(* IEC 61131-3 sources: daoli-st-library/DL_MathData (part 12) *)

(* ---- FC_DL_DintMsToTod.st ---- *)
(*
    FC_DL_DintMsToTod —— 当日毫秒到 TOD 的防御转换
    ------------------------------------------------------------------
    分类      : DL_MathData / TimeConv
    前缀      : FC_DL_
    版本      : 1.0.0
    溯源      : IEC 61131-3 标准 TOD 语义的道莅防御性实现；本件为
                FC_DL_TodToDintMs 的严格逆运算，接口语义由标准定义，
                内部委托平台内建 DINT_TO_TOD，不自行按时基重算；
                外围错误分级、单圈折回、双端钳位与双语文档 100% 自有；
                clean-room 重写，未复制任何闭源厂商源码，参考实现仅限 MIT/Apache 许可
    平台      : 纯 IEC 61131-3，CODESYS V3.5+ / TwinCAT 3 / InoProShop 通用
    作者      : 道莅代码库 · PLC编程专家（R19）
    ------------------------------------------------------------------
    功能说明  : 把「自当日 00:00 起的毫秒数」还原为 TOD，供上层排程件与定时器比较。
                有效域 0~86399999 ms；可接受域 -86400000~172799999 ms（含跨日正负各一圈）。
                核心防御：① 超可接受域直接故障级 031E 早退，绝不对非法值调内建；
                ② 负值按单圈折回当日（先判后算，仅一圈内成立，无循环语句）；
                ③ 钳位只在 0 与 86399999 ms 两端，越界量由 bClampSilently 决定分级；
                ④ 交付门槛：委托 DINT_TO_TOD 内建链，须在 CODESYS / TwinCAT 3 /
                   InoProShop 三平台各编译验证一次（跨平台时间类转换链行为存疑）。
                职责边界：本件只做数值还原，不判时区、不做日历进位。
    错误码    : 16#0001_0400 输入越当日域已被钳位到 0 或 86399999 ms——信息级，正常防御
                16#0001_0401 预留禁用（信息级，不得挪用）
                16#0001_031E 输入超可接受域（< -86400000 ms 或 > 172799999 ms）——故障级，返回 T#0S 且 bValid = FALSE
                16#0001_031F 调用方要求不静默（bClampSilently = FALSE）且发生钳位——故障级，返回钳位值但 bValid = FALSE
                16#0001_0320 预留禁用（故障级，不得挪用）
    码位总账  : 16#0001_0400 用 / 16#0001_0401 预留 ｜ 16#0001_031E 用 / 16#0001_031F 用 / 16#0001_0320 预留
    状态机    : R6 标注 N/A —— 本组件为纯函数无顺序状态机，无 CASE 可写，非法状态不可能出现
    采样约定  : 本件无定时器、无沿检测、无顺序状态；单拍纯计算，结论与任务周期无关。
    修订记录  : 2026-11-16 v1.0.0 首次入库（R19）
*)
FUNCTION FC_DL_DintMsToTod : TOD
VAR_INPUT
    nMsOfDay        : DINT := 0;              // 当日毫秒偏移 [ms]，有效域 0~86399999，可接受域 -86400000~172799999 / day-millisecond offset [ms], valid 0~86399999, accepted -86400000~172799999
    bClampSilently  : BOOL := TRUE;           // TRUE = 越界钳位只置信息码；FALSE = 越界置故障级 / TRUE clamps with info code only, FALSE raises a fault level
END_VAR
VAR_OUTPUT
    eErr            : UDINT;                  // 错误码，0=正常 / error id, 0=ok
    bError          : BOOL;                   // 故障标志，eErr 为故障级时 TRUE / error flag, TRUE on fault-level eErr
    bValid          : BOOL;                   // 返回值是否可用 / return value valid flag
    bClamped        : BOOL;                   // 本拍是否发生钳位 / clamp event in this cycle
END_VAR
VAR CONSTANT
    DL_TOD_MS_MIN   : DINT := 0;              // 当日毫秒下界 [ms] / day-millisecond lower bound [ms]
    DL_TOD_MS_MAX   : DINT := 86399999;       // 当日毫秒上界（24 h − 1 ms） [ms] / day-millisecond upper bound, 24 h minus 1 ms [ms]
    DL_TOD_DAY_MS   : DINT := 86400000;       // 一整天毫秒数（单圈折回用） [ms] / milliseconds of one day, for single-wrap folding [ms]
    DL_TOD_MS_MIN_EXT : DINT := -86400000;    // 可接受下界（跨日回退一圈） [ms] / accepted lower bound, one day backwards [ms]
    DL_TOD_MS_MAX_EXT : DINT := 172799999;    // 可接受上界（跨日超前一圈） [ms] / accepted upper bound, one day forwards [ms]
END_VAR
VAR
    nMs             : DINT;                   // 折回与钳位后的中间毫秒值 [ms] / intermediate millisecond value after folding and clamping [ms]
END_VAR

// 段 1｜返回值与错误状态预置 / segment 1, preset return value and error status
FC_DL_DintMsToTod := T#0S;                    // 故障缺省返回当日零点 / fault default returns midnight
eErr := 0;                                    // 预置无错误 / preset no error
bError := FALSE;                              // 预置无故障 / preset no fault
bValid := FALSE;                              // 预置不可用，通过闸门后置位 / preset invalid, set TRUE after the gates
bClamped := FALSE;                            // 预置未钳位 / preset no clamp

// 段 2｜可接受域闸门（越一圈直接故障级，绝不对非法值调内建）/ segment 2, accepted domain gate
IF (nMsOfDay < DL_TOD_MS_MIN_EXT) OR (nMsOfDay > DL_TOD_MS_MAX_EXT) THEN
    eErr := 16#0001_031E;                     // 超可接受域故障码 / accepted domain exceeded fault id
    bError := TRUE;                           // 置故障标志 / raise the error flag
    bValid := FALSE;                          // 返回值不可用 / return value not usable
    FC_DL_DintMsToTod := T#0S;                // 明确返回零点，不用非法值调内建 / return midnight explicitly, never feed an illegal value to the built-in
    RETURN;                                   // 故障级提前返回 / early return on fault
END_IF

// 段 3｜负值单圈折回当日（先判后算，无循环语句）/ segment 3, fold negative values back by one day
nMs := nMsOfDay;                              // 取入参副本参与运算，不改调用方数据 / copy the input, never modify caller data
IF nMs < DL_TOD_MS_MIN THEN
    nMs := nMs + DL_TOD_DAY_MS;               // 单圈折回：域已由段 2 保证 |nMs| ≤ 一圈 / single wrap is enough, segment 2 bounded the magnitude to one day
END_IF

// 段 4｜当日双端钳位（永不对非法值直接调内建）/ segment 4, clamp on both day bounds
IF nMs < DL_TOD_MS_MIN THEN
    nMs := DL_TOD_MS_MIN;                     // 防御性兜底：折回后仍为负则钳 0 ms / defensive floor, clamp to 0 ms if still negative
    bClamped := TRUE;                         // 记录钳位事件 / record the clamp event
ELSIF nMs > DL_TOD_MS_MAX THEN
    nMs := DL_TOD_MS_MAX;                     // 越上界钳 86399999 ms（24 h − 1 ms） / clamp to 86399999 ms, 24 h minus 1 ms
    bClamped := TRUE;                         // 记录钳位事件 / record the clamp event
END_IF

// 段 5｜钳位分级：静默只置信息码，不静默置故障级但返回钳位值 / segment 5, clamp severity
IF bClamped THEN
    IF bClampSilently THEN
        eErr := 16#0001_0400;                 // 信息级：越当日域已钳位，正常防御，不置故障 / info level, clamped into the day domain, no fault raised
        bValid := TRUE;                       // 钳位值仍可用 / the clamped value is usable
    ELSE
        eErr := 16#0001_031F;                 // 故障级：调用方要求不静默 / fault level, the caller refused silent clamping
        bError := TRUE;                       // 置故障标志 / raise the error flag
        bValid := FALSE;                      // 钳位结果标记为不可用 / the clamped result is flagged unusable
    END_IF
ELSE
    eErr := 0;                                // 一轮内合法输入不进钳位分支 / in-domain input never enters the clamp branch
    bValid := TRUE;                           // 域内结果可用 / in-domain result is usable
END_IF

// 段 6｜委托内建转换（入参已保证落在 0~86399999 ms）/ segment 6, delegate to the built-in conversion
FC_DL_DintMsToTod := DINT_TO_TOD(nMs);        // 委托内建，不自行按时基累加 / delegate to the built-in, never accumulate the time base by hand
END_FUNCTION

(* ---- FC_DL_DintToBcd.st ---- *)
(*
  ==================================================================
  组件名 Component  : FC_DL_DintToBcd
  分类   Category   : DL_MathData
  前缀   Naming     : FC_DL_ ｜ b/n/u/f/t/e/st 类型前缀制（R265）
  码位   Code ID    : 16#0001_0658（故障级）
  版本   Version    : 1.0.0
  复杂度 Complexity  : 低
  功能   Purpose    : DINT → 8 位 BCD（DWORD 容器），负值显式拒绝 + 越域显式拒绝，
                      逐位 MOD 10 / DIV 10 提取后按权装入半字节。
  开源溯源 Origin    : 公开公式 clean-room，参考 BCD 编码公开工程语义（分类与参数域
                      借鉴，零代码复制），本件实现、闸门与码位 100% 自有。
  许可证 License    : MIT
  参考   Reference  : IEC 61131-3:2013 §6.6 算术与移位运算符（MOD / DIV / SHL / OR）
  平台   Platform   : 纯 IEC 61131-3（FOR / MOD / DIV / SHL / OR），三平台通用
  依赖   Depends    : 仅 Standard.library（无库调用）
  分工声明 Split     : FC_DL_ByteToBcd / FC_DL_WordToBcd / FC_DL_UdintToBcd 为既有
                      BCD 编码族（无符号域入口），本件为 DINT 带符号域入口；负值
                      显式拒绝为本件与 UDINT 版本的**行为差异**（写死，禁取绝对值
                      回绕伪装成功）；MOD/DIV 10 原语经派单规格明写授权，本件为
                      BCD 编解码属主；四件互引（R216）。
  归属 Ownership     : 本件无 TYPE 声明；全部引脚为 IEC 标准原生类型。
  ------------------------------------------------------------------
  边界 Boundary     :
                      一 判据顺序（写死）：① nIn < 0 → 故障级码 + udBcd = 0 早退
                         （负值不可 BCD 表示，禁取绝对值回绕）；② nIn > 99999999 →
                         越域故障 + bOvF = TRUE 早退；③ 正常才进入提取；
                      二 两场景一码的反证句（R90）：负值与越域的出口仅 bOvF 一位
                         之差（负值 FALSE / 越域 TRUE），一个输出位即可唯一还原
                         场景，三组以内输出可区分，按 R90 不另立码；
                      三 移位量 4·k（k = 0..7）最大 28 < 32（DWORD 位宽），结构性
                         安全（R48）；
                      四 越域上界常量 DL_BCD_MAX = 99999999 与 8 位 BCD 可表域
                         一致，超域属「不可表」而非「截断后仍可用」，禁静默截断；
                      五 纯函数：无记忆量、无定时器、无边沿实例，每调用重算；
                      六 无全局、无外部变量、无物理地址、无指针。
  错误码 Codes      :
    16#0001_0658【故障级】不可 BCD 编码（nIn < 0 负值，bOvF = FALSE；或
                         nIn > 99999999 越域，bOvF = TRUE）
  码位反证 Note     :
    负值与越域共用一码：出口组合仅 bOvF 一位可区分（边界二反证句），按 R90 不另立。
  验收 Acceptance   :
    算法已证（脚本）：未跑 ｜ 编译器已证（三平台）：未跑
    V1 0 → 16#00000000；V2 99999999 → 16#99999999（恰好整除上界向量）
    V3 -1 → 故障 0658 + bOvF = FALSE + 早退（禁取绝对值）
    V4 100000000 → 故障 0658 + bOvF = TRUE + 早退
    V5 12345678 → 16#12345678
  修订记录 Revision  :
    2026-11-21  v1.0.0  R63 首版（批 1 · 序号 2）
  ==================================================================
*)
FUNCTION FC_DL_DintToBcd : BOOL
VAR_INPUT
    nIn     : DINT := 0; // 待编码整数 [个]，合法域 0..99999999 / the integer to encode, legal from zero to ninety nine million
END_VAR
VAR_OUTPUT
    udBcd   : DWORD := 16#00000000; // 8 位 BCD 输出 [码] / the eight digit BCD output
    bOvF    : BOOL := FALSE;        // 越域标志（仅 nIn > 99999999 置位）[-] / the overflow flag raised only above the BCD domain
    bValid  : BOOL := FALSE;        // 结果可用 [-] / the result usable flag
    eErr    : UDINT := 16#0000_0000; // 错误码，0 = 正常 / the error code, zero is ok
    bError  : BOOL := FALSE;        // 故障标志（故障级码同拍置位，R45 配对）/ the fault flag raised with a fault level code
END_VAR
VAR
    k       : DINT := 0;  // 码元位置索引 [下标]，0..7 / the digit position index from zero to seven
    nShift  : DINT := 0;  // 移位量 [位]，4·k ≤ 28 结构性安全 / the shift amount of four times the position, proven below the word width
    nWork   : DINT := 0;  // 逐位提取工作副本 [个] / the working copy of the digit extraction
    uDig    : USINT := 0; // 当前位码元 [位] / the current digit extracted
END_VAR  // R64 结构补齐：VAR 段缺失的 END_VAR（门禁机械修复）
VAR CONSTANT
    DL_BCD_MAX   : DINT := 99999999;   // 8 位 BCD 可表上界 [个] / the representable ceiling of the eight digit BCD
    DL_BCD_N     : DINT := 8;          // 码元总数 [个] / the digit count of eight
    DL_BCD_TEN   : DINT := 10;         // 十进制提取基数 [个] / the decimal extraction base of ten
    DL_BCD_NIB   : DINT := 4;          // 每码元位宽 [位] / the nibble width of four bits
    DL_BCD_ZERO  : DINT := 0;          // 整型零常量 [个] / the integer zero constant
    DL_BCD_ONE   : DINT := 1;          // 整型一常量 [个] / the integer one constant
END_VAR

// 段 1｜返回值与全部出口预置安全值（R45 四段式第一段）/ segment 1, the preset of the return and every outlet
FC_DL_DintToBcd := FALSE; // 返回值预置假 / preset the return false
udBcd := 16#00000000; // BCD 输出预置全零 [码] / preset the BCD output to all zeros
bOvF := FALSE; // 越域标志预置假 / preset the overflow flag false
bValid := FALSE; // 可用标志预置假 / preset the validity false
eErr := 16#0000_0000; // 错误码预置正常 / preset the code to ok
bError := FALSE; // 故障标志预置假 / preset the error flag false
nWork := DL_BCD_ZERO; // 工作副本预置零 [个] / preset the working copy zero
k := DL_BCD_ZERO; // 索引预置零 / preset the index zero
nShift := DL_BCD_ZERO; // 移位量预置零 [位] / preset the shift amount zero
uDig := 0; // 码元预置零 [位] / preset the digit zero

// 段 2｜判据一：负值显式拒绝（边界一①，禁取绝对值回绕伪装成功）/ segment 2, the negative value rejection
IF nIn < DL_BCD_ZERO THEN // 负值不可 BCD 表示 / a negative value is not representable in BCD
    udBcd := 16#00000000; // 输出强制全零 [码] / force the output to all zeros
    eErr := 16#0001_0658; // 故障级：不可 BCD 编码（负值，bOvF 保持 FALSE 供区分）/ fault grade, not encodable as BCD, the overflow flag stays false for the discrimination
    bError := TRUE; // 同拍置故障标志（R45 配对）/ raise the fault flag on the same scan
    bValid := FALSE; // 结果不可用 / the result is not usable
    RETURN; // 早退 / early return
END_IF

// 段 3｜判据二：越域显式拒绝（边界一②，禁静默截断）/ segment 3, the domain overflow rejection
IF nIn > DL_BCD_MAX THEN // 超 8 位 BCD 可表上界 / above the representable ceiling
    udBcd := 16#00000000; // 输出强制全零 [码] / force the output to all zeros
    bOvF := TRUE; // 置越域标志（与负值场景的唯一区分位）/ raise the overflow flag, the only bit distinguishing this scene
    eErr := 16#0001_0658; // 故障级：不可 BCD 编码（越域）/ fault grade, not encodable as BCD, the domain is exceeded
    bError := TRUE; // 同拍置故障标志（R45 配对）/ raise the fault flag on the same scan
    bValid := FALSE; // 结果不可用 / the result is not usable
    RETURN; // 早退 / early return
END_IF

// 段 4｜逐位提取与按权装入（移位量 4·k ≤ 28 < 32 结构性安全，边界三）/ segment 4, the digit extraction and the weighted packing
nWork := nIn; // 工作副本接管 [个] / take the working copy
FOR k := DL_BCD_ZERO TO DL_BCD_N - DL_BCD_ONE DO // 有界遍历 8 个码元位置 / the bounded traversal over eight digit positions
    uDig := DINT_TO_USINT(nWork MOD DL_BCD_TEN); // 当前位 = nWork MOD 10 [位] / the current digit is the remainder of ten
    nWork := nWork / DL_BCD_TEN; // 副本右移一位（DINT 整除截断，nIn ≥ 0 已证，无负回绕）/ shift the copy one digit right, the truncating division is safe since the input is proven non negative
    nShift := DL_BCD_NIB * k; // 移位量 = 4·k，最大 28 [位] / the shift amount of four times the position
    udBcd := udBcd OR SHL(USINT_TO_DWORD(uDig), nShift); // 码元装入对应半字节（OR 合成）/ pack the digit into its nibble by the or composition
END_FOR

// 段 5｜统一出口 / segment 5, the unified outlet
bValid := TRUE; // 结果可用 / the result is usable
FC_DL_DintToBcd := TRUE; // 返回成功 / return success
END_FUNCTION

(* ---- FC_DL_DintToRealChk.st ---- *)
(*
    FC_DL_DintToRealChk —— DINT 到 REAL 精度告警转换
    ------------------------------------------------------------------
    分类      : DL_MathData / Convert
    前缀      : FC_DL_
    版本      : 1.0.0
    溯源      : IEC 61131-3 标准语义的道莅防御性实现
                （接口语义由 IEC 61131-3 定义，内部委托平台内建 DINT_TO_REAL，
                  外围统一错误码 / 钳位 / 双语文档；clean-room 重写，
                  未复制任何闭源厂商源码，参考实现仅限 MIT/Apache 许可）
    平台      : 纯 IEC 61131-3，CODESYS / TwinCAT / InoProShop 通用
    作者      : 道莅代码库 · PLC编程专家（R17）
    ------------------------------------------------------------------
    功能说明  : 将 DINT 防御性转换为 REAL 并作为返回值输出，转换委托平台内建 DINT_TO_REAL；
                |nIn| 超过 2^24（16777216，REAL 尾数 24 位可精确表示的整数上界）时，
                值照常转换输出，仅置信息级 16#0001_01FC 提示低位精度损失（bError=FALSE、bValid=TRUE）；
                极值对称性防御：采用双侧比较 nIn > 上界 OR nIn < -上界，
                禁用 ABS(nIn) 单侧比较（对 DINT 最小值无回绕，但保持与 R16 LintToLrealChk 同范式，避免后续升位改造引入回绕）；
                钳位方向：无钳位（信息级仅记录，转换结果为最接近的可表值）。
    错误码    : 16#0001_01FC |nIn| 超 2^24 精度极限，转换值低位可能失真——信息级，正常防御
                16#0001_01FD 预留禁用（信息级，不得挪用）
                16#0001_02E8 预留禁用（故障级，不得挪用）
                16#0001_02E9 预留禁用（故障级，不得挪用）
                16#0001_02EA 预留禁用（故障级，不得挪用）
    状态机    : R6 标注 N/A —— 本组件为纯函数无顺序状态机，无 CASE 可写，非法状态不可能出现，故以本节说明替代 ELSE 兜底
    修订记录  : 2026-11-16 v1.0.0 首次入库（R17）
*)
FUNCTION FC_DL_DintToRealChk : REAL
VAR_INPUT
    nIn : DINT; // 待转换整数值，建议域 ±2147483647 [无量纲] / integer value to convert, suggested domain +/-2147483647 [dimensionless]
END_VAR
VAR_OUTPUT
    eErr   : UDINT; // 错误码，0=正常 / error id, 0=ok
    bError : BOOL;  // 是否出错，eErr 非 0 时为 TRUE / error flag, TRUE when eErr is nonzero
    bValid : BOOL;  // 输出是否有效可用 / output valid flag
END_VAR
VAR CONSTANT
    DL_F24_MAX : DINT := 16777216; // REAL 尾数 24 位可精确表示的整数上界 2^24 [无量纲] / 2^24 exact-integer bound of REAL's 24-bit significand [dimensionless]
    DL_REAL_ZERO : REAL := 0.0;    // 返回值预置零（本件无故障路径，仅作预置约定） [无量纲] / preset zero, no fault path in this component [dimensionless]
END_VAR

// 段 1｜返回值与错误状态预置 / segment 1, preset return value and error status
FC_DL_DintToRealChk := DL_REAL_ZERO; // 预置 0.0（本件无故障级路径，仅作预置约定） [无量纲] / preset 0.0, no fault-level path in this component [dimensionless]
eErr   := 0;     // 预置无错误 / preset no error
bError := FALSE; // 预置无故障（本件无故障级路径） / preset no fault, no fault-level path here
bValid := FALSE; // 预置输出无效，通过精度判定后置位 / preset invalid, set TRUE after the precision check

// 段 2｜24 位尾数精度极限判定与主体转换（末段） / segment 2, 24-bit significand precision check and main conversion (final)
FC_DL_DintToRealChk := DINT_TO_REAL(nIn); // 值照常转换（委托平台内建转换语义），本件只告警不钳位 [无量纲] / convert as-is via the built-in conversion, this component warns but never clamps [dimensionless]
IF (nIn > DL_F24_MAX) OR (nIn < -DL_F24_MAX) THEN // 双侧比较，禁用 ABS 单侧式 [无量纲] / two-sided comparison, single-sided ABS form forbidden [dimensionless]
    eErr := 16#0001_01FC; // 信息级：超 2^24 精度极限，低位可能失真，仅记录不钳位 / info level: beyond the 2^24 precision limit, low bits may lose accuracy, recorded only
ELSE
    eErr := 0;            // 精度域内无告警 / within the precision domain, no notice
END_IF
bError := FALSE; // 信息级精度告警不置故障 / info-level precision notice never raises fault
bValid := TRUE;  // 域内或精度告警输出均有效可用 / in-domain or precision-noticed output is valid
END_FUNCTION

(* ---- FC_DL_DintToStringTrim.st ---- *)
(*
    FC_DL_DintToStringTrim —— DINT 到 STRING 的防御字符串化
    ------------------------------------------------------------------
    分类      : DL_MathData / Convert
    前缀      : FC_DL_
    版本      : 1.0.0
    溯源      : IEC 61131-3 标准语义的道莅防御性实现（DINT → STRING，去前导空格与长度钳位）；
                委托平台内建 DINT_TO_STRING 与标准串函数 LEN / MID / LEFT，本件不重实现格式化内核；
                空格修剪、四步截断样板、目标长度闸、错误分级与码位 100% 自有；
                clean-room 重写，未复制任何闭源厂商源码，参考实现仅限 MIT/Apache 许可
    平台      : 纯 IEC 61131-3，CODESYS V3.5+ / TwinCAT 3 / InoProShop 通用
    作者      : 道莅代码库 · PLC编程专家（R20）
    ------------------------------------------------------------------
    功能说明  : 数值要拼进 CSV 行、报文帧、条码内容、文件名时，必须先字符串化。
                各平台 DINT_TO_STRING 的右对齐习惯不一：有的前置空格补齐到固定宽度，
                有的不留空格。带空格的数值混进 CSV 会多出一列，拼进报文会错位一个字节，
                而这类故障在 PLC 侧完全静默，只有上位机解析时才暴露。
                核心防御：① 逐字符定位首个非空格后一次 MID 截取，杜绝「逐字符拼串」的
                   长度与性能问题（拼串会随长度平方级增长）。
                ② 扫描用定长 FOR（上界 255），禁用 WHILE——串函数异常时 WHILE 会死循环，
                   FOR 上界结构性封顶。
                ③ 截断走四步样板（R37）：先把长度一次锁存 → 与目标宽度比较 →
                   截断标志置位先于任何写入 → 按 bAllowTrunc 分路；不允许截断时返回空串
                   并升故障级，绝不返回半截数值——半截数值形如把 12345 写成 123，
                   上位机会把它当成真实数据。
                ④ uTargetMax 引脚钳位在 1~255：0 长度目标无意义；255 是 STRING 型上限（R49 口径），
                   USINT 类型本身的 255 上界即为其第二道保险。
                职责边界：LREAL 字符串化（含非有限值统一文本）归 FC_DL_LrealToStringTrim；
                串处理九函数归 T0-6 家族；本件只管整型方向。
    编译门槛  : 主路径依赖平台内建 DINT_TO_STRING 与标准串函数 LEN / MID / LEFT。
                DINT_TO_STRING 的返回宽度平台间不同（有 11 字符起的多种取值），
                故本件不假设其宽度，一律按 LEN 实测后处理，必要时再按目标长度钳位。
    错误码    : 16#0001_0426 已修剪前导空格（bTrimmed 可查）——信息级，值可用
                16#0001_0427 发生截断且 bAllowTrunc = TRUE（bTruncated 可查）——信息级，值可用
                16#0001_0357 目标长度非法（uTargetMax = 0，或平台 USINT 上限异常）——故障级，返回空串
                16#0001_0358 需要截断但 bAllowTrunc = FALSE——故障级，返回空串
                16#0001_0359 预留禁用（故障级，不得挪用）
    码位总账  : 16#0001_0426 用 / 16#0001_0427 用 ｜ 16#0001_0357 用 / 16#0001_0358 用 / 16#0001_0359 预留
    状态机    : R6 标注 N/A —— 本组件为纯函数无顺序状态机，无 CASE 可写，非法状态不可能出现
    采样约定  : 本件无定时器、无沿检测、无状态；单拍纯计算，结论与任务周期无关。
    修订记录  : 2026-11-16 v1.0.0 首次入库（R20）
*)
FUNCTION FC_DL_DintToStringTrim : STRING(255)
VAR_INPUT
    nIn              : DINT;                  // 待字符串化的数值 [无量纲]，全域 / value to serialise [dimensionless], full DINT domain
    uTargetMax       : USINT := 31;           // 目标缓冲可用长度 [字符]，1~255 / usable target length [characters], 1 to 255
    bAllowTrunc      : BOOL := FALSE;         // TRUE = 允许截断；FALSE = 需截断即故障 / TRUE allows truncation, FALSE turns it into a fault
END_VAR
VAR_OUTPUT
    eErr             : UDINT;                 // 错误码，0=正常 / error id, 0=ok
    bError           : BOOL;                  // 故障标志，eErr 为故障级时 TRUE / error flag, TRUE on fault-level eErr
    bValid           : BOOL;                  // 返回值是否可用（故障级为 FALSE）/ return usable, FALSE on fault level
    bTrimmed         : BOOL;                  // 修剪了前导空格 / leading blanks were trimmed
    bTruncated       : BOOL;                  // 超目标长度发生截断 / truncation to the target length happened
END_VAR
VAR CONSTANT
    DL_STR_CAP_MAX   : USINT := 255;          // STRING 型长度上限 [字符]，R49 口径 / STRING capacity [characters], per R49
    DL_STR_TARGET_MIN : USINT := 1;           // 目标长度下限 [字符] / target length lower bound [characters]
    DL_STR_SCAN_MAX  : INT := 255;            // 扫描上界 [字符]，与 STRING 上限一致 / scan bound [characters], equals the STRING capacity
    DL_STR_BLANK     : STRING(1) := ' ';      // 单个空格字符，修剪判据 / a single blank used by the trim test
    DL_STR_EMPTY     : STRING(1) := '';       // 空串常量，故障缺省返回 / empty string returned on faults
    DL_INT_ZERO      : INT := 0;              // 整型零常量，避免裸字面量 [字符] / integer zero constant [characters]
    DL_INT_ONE       : INT := 1;              // 整型一常量，首个非空格位置起点 [字符] / integer one constant, first non-blank position [characters]
END_VAR
VAR
    sRaw             : STRING(255);           // 内建字符串化原始结果 / raw result of the built-in conversion
    sTrim            : STRING(255);           // 修剪后的中间串 / intermediate string after the trim
    sOut             : STRING(255);           // 最终输出串 / final output string
    nLen             : INT;                   // 原始串有效长度 [字符] / effective length of the raw string [characters]
    nStart           : INT;                   // 首个非空格位置，1 起始，0 = 全为空格 / first non-blank position, 1-based, 0 means all blanks
    nIdx             : INT;                   // 扫描游标 [字符]，1 起始 / scan cursor [characters], 1-based
    nKept            : INT;                   // 修剪后保留长度，一次锁存 [字符] / retained length, latched exactly once [characters]
    nTarget          : INT;                   // 目标长度，由引脚转出 [字符] / target length derived from the pin [characters]
    bFound           : BOOL;                  // 已找到首个非空格标志 / a first non-blank has been found
END_VAR

// 段 1｜返回值与错误状态预置 / segment 1, preset return value and error status
FC_DL_DintToStringTrim := DL_STR_EMPTY;       // 故障缺省返回空串 / fault default returns an empty string
eErr := 0;                                    // 预置无错误 / preset no error
bError := FALSE;                              // 预置无故障 / preset no fault
bValid := FALSE;                              // 预置不可用，通过闸门后置位 / preset invalid, set TRUE after the gates
bTrimmed := FALSE;                            // 预置未修剪 / preset no trim
bTruncated := FALSE;                          // 预置未截断 / preset no truncation
sOut := DL_STR_EMPTY;                         // 输出串清零 / clear the output string
nKept := DL_INT_ZERO;                         // 保留长度清零 / clear the retained length

// 段 2｜目标长度闸：0 长度目标无意义，先判后算 / segment 2, target length gate
IF uTargetMax < DL_STR_TARGET_MIN THEN
    eErr := 16#0001_0357;                     // 故障级：目标长度非法，返回空串 / fault level, illegal target length, return an empty string
    bError := TRUE;                           // 置故障标志 / raise the error flag
    bValid := FALSE;                          // 返回值不可用 / flag the return as unusable
    RETURN;                                   // 出口，不触碰内建 / exit, the built-in is never touched
END_IF
nTarget := USINT_TO_INT(uTargetMax);          // 目标长度转整型 [字符] / convert the target length into an integer [characters]
IF nTarget > USINT_TO_INT(DL_STR_CAP_MAX) THEN
    nTarget := USINT_TO_INT(DL_STR_CAP_MAX);  // 双保险：按 STRING 上限钳位 [字符] / second line of defence, clamp to the STRING capacity [characters]
END_IF

// 段 3｜主体：委托平台内建字符串化 / segment 3, delegate the built-in conversion
sRaw := DINT_TO_STRING(nIn);                  // 数值 → 原始串（可能含前导空格）/ value to raw string, possibly blank padded

// 段 4｜有效长度一次锁存并钳位 / segment 4, latch the effective length once and clamp it
nLen := LEN(sRaw);                            // 原始串长度 [字符] / raw string length [characters]
IF nLen > DL_STR_SCAN_MAX THEN
    nLen := DL_STR_SCAN_MAX;                  // 超容量按上限钳位 [字符] / clamp to the capacity [characters]
ELSIF nLen < DL_INT_ZERO THEN
    nLen := DL_INT_ZERO;                      // 负长度防御，结构性不可达 [字符] / negative length guard, structurally unreachable [characters]
END_IF

// 段 5｜前导空格修剪：定长 FOR 扫描，禁 WHILE / segment 5, leading blank trim with a bounded FOR loop
nStart := DL_INT_ZERO;                        // 0 表示尚未找到非空格 / zero means no non-blank found yet
bFound := FALSE;                              // 扫描标志预置 / preset the scan flag
FOR nIdx := DL_INT_ONE TO nLen DO
    IF NOT bFound THEN
        IF MID(sRaw, DL_INT_ONE, nIdx) <> DL_STR_BLANK THEN
            nStart := nIdx;                   // 记录首个非空格位置 [字符] / record the first non-blank position [characters]
            bFound := TRUE;                   // 扫描标志置位 / raise the scan flag
        END_IF
    END_IF
END_FOR

IF nStart = DL_INT_ZERO THEN
    sTrim := DL_STR_EMPTY;                    // 全为空格：合法的空结果，不是错误 / all blanks, a legal empty result
ELSE
    sTrim := MID(sRaw, nLen - nStart + DL_INT_ONE, nStart); // 一次截取中间段 / extract the retained segment in one call
    IF nStart > DL_INT_ONE THEN
        bTrimmed := TRUE;                     // 确实修剪了前导空格 / blanks were really trimmed
        eErr := 16#0001_0426;                 // 信息级：已修剪前导空格 / info level, leading blanks were trimmed
    END_IF
END_IF

// 段 6｜四步截断样板（R37）：长度锁存 → 宽度比较 → 标志先置 → 按允许分路 / segment 6, the four-step truncation pattern
nKept := LEN(sTrim);                          // 修剪后长度，一次锁存 [字符] / retained length, latched once [characters]
IF nKept > nTarget THEN
    bTruncated := TRUE;                       // 标志先于任何写入 / the flag precedes every write
    IF bAllowTrunc THEN
        sOut := LEFT(sTrim, nTarget);         // 允许截断：按目标长度截取 / truncation allowed, take the target length
        eErr := 16#0001_0427;                 // 信息级：发生截断，值可用 / info level, truncated, still usable
    ELSE
        eErr := 16#0001_0358;                 // 故障级：需截断但不允许 / fault level, truncation needed but not allowed
        bError := TRUE;                       // 置故障标志 / raise the error flag
        bValid := FALSE;                      // 返回值不可用 / flag the return as unusable
        FC_DL_DintToStringTrim := DL_STR_EMPTY; // 返回空串，绝不返回半截数值 / return an empty string, never a partial number
        RETURN;                               // 出口 / exit
    END_IF
ELSE
    sOut := sTrim;                            // 无需截断，直接采用修剪结果 / no truncation, take the trimmed string
END_IF

// 段 7｜发布结果 / segment 7, publish the result
FC_DL_DintToStringTrim := sOut;               // 输出最终串 / publish the final string
bValid := TRUE;                               // 修剪/截断/直通均可用 / usable in every published path
bError := FALSE;                              // 信息级不置故障（双保险）/ info level never raises a fault, second line of defence
END_FUNCTION

(* ---- FC_DL_DintToUintSat.st ---- *)
(*
    FC_DL_DintToUintSat —— DINT 到 UINT 饱和防御转换
    ------------------------------------------------------------------
    分类      : DL_MathData / Convert
    前缀      : FC_DL_
    版本      : 1.0.0
    溯源      : IEC 61131-3 标准语义的道莅防御性实现
                （内部委托平台内建函数，外围统一错误码/钳位/双语文档；
                  未复制任何闭源厂商源码，参考实现仅限 MIT/Apache 许可）
    平台      : 纯 IEC 61131-3，CODESYS / TwinCAT / InoProShop 通用
    作者      : 道莅代码库 · PLC编程专家（R16）
    ------------------------------------------------------------------
    功能说明  : 将 DINT 输入防御性转换为 UINT 并作为返回值输出；
                nIn < 0 时钳位至 0，置信息级 16#0001_01CA（UINT 无符号，负值不可表）；
                nIn 超出 UINT 上界 65535 时钳位至上界，置信息级 16#0001_01CB；
                钳位方向：下界 0 / 上界 65535（双侧饱和）；
                纯整数域输入不存在 NaN/±INF 非有限态，亦无除法运算，故本组件无故障级路径；
                域内转换委托平台内建 DINT_TO_UINT 语义，不重实现数学内核；
                信息级码属正常防御：bError=FALSE、bValid=TRUE，输出钳位后防御值。
    错误码    : 16#0001_01CA 负值输入，已钳位至 0——信息级，正常防御
                16#0001_01CB 输入超 UINT 上界，已钳位至 65535——信息级，正常防御
                16#0001_029D 预留禁用（故障级，不得挪用）
                16#0001_029E 预留禁用（故障级，不得挪用）
                16#0001_029F 预留禁用（故障级，不得挪用）
    状态机    : R6 标注 N/A —— 本组件为纯函数无顺序状态机，无 CASE 可写，非法状态不可能出现，故以本节说明替代 ELSE 兜底
    修订记录  : 2026-11-16 v1.0.0 首次入库（R16）
*)
FUNCTION FC_DL_DintToUintSat : UINT
VAR_INPUT
    nIn : DINT; // 待转换输入 [无量纲] / input value to convert
END_VAR
VAR_OUTPUT
    eErr   : UDINT; // 错误码，0=正常 / error id, 0=ok
    bError : BOOL;  // 是否出错，eErr 非 0 时为 TRUE / error flag, TRUE when eErr is nonzero
    bValid : BOOL;  // 输出是否有效可用 / output valid flag
END_VAR
VAR CONSTANT
    DL_UINT16_MAX : DINT := 65535; // UINT 域上界 65535 [无量纲] / UINT upper bound 65535
END_VAR

// 段 1｜返回值与错误状态预置 / segment 1, preset return value and error status
FC_DL_DintToUintSat := 0; // 故障缺省返回 0 [无量纲] / fault default returns 0
eErr   := 0;     // 预置无错误 / preset no error
bError := FALSE; // 预置无故障（整数域无故障态） / preset no fault (no fault states in integer domain)
bValid := FALSE; // 预置无效，通过钳位判定后置位 / preset invalid, set TRUE after clamp check

// 段 2｜双侧饱和钳位与主体转换（末段） / segment 2, double-side saturating clamp and main conversion (final)
IF nIn < 0 THEN
    FC_DL_DintToUintSat := 0; // 负值钳位至 0（UINT 无符号语义） / negative input clamped to 0 (UINT is unsigned)
    eErr := 16#0001_01CA;     // 信息级：负值已钳零 / info level: negative input clamped to zero
ELSIF nIn > DL_UINT16_MAX THEN
    FC_DL_DintToUintSat := 16#FFFF; // 正向钳位至 UINT 上界 65535 / clamp to UINT upper bound 65535
    eErr := 16#0001_01CB;           // 信息级：超上界已钳位 / info level: above upper bound, clamped
ELSE
    FC_DL_DintToUintSat := DINT_TO_UINT(nIn); // 域内委托平台内建 _TO_ 转换语义 / in-domain delegate to built-in _TO_ conversion
    eErr := 0; // 域内无错误 / in-domain, no error
END_IF
bValid := TRUE; // 域内或钳位输出均有效可用 / in-domain or clamped output is valid
END_FUNCTION

(* ---- FC_DL_DivDintSafeChk.st ---- *)
(*==============================================================================
 * 组件名称 (Component)  : FC_DL_DivDintSafeChk
 * 所属子库 (Sublibrary) : DL_MathData
 * 归属目录 (Directory)  : C:\Library\DL_MathData
 * 当前版本 (Version)    : 1.0.0
 * 分类/来源标签         : 函数（FUNCTION）· 纯函数 · DINT 安全除
 *                         iec-std-wrapper / math-safe
 * 兼容性   (Platform)   : CODESYS 3.5 / TwinCAT 3 / 汇川 InoProShop / 施耐德
 *                         Machine Expert；仅用 IEC 标准 DINT 除法与 MOD 语义
 * 溯源声明 (Provenance) : IEC 61131-3 标准语义的道莅防御性实现——内部委托平台标准库语义，
 *                         外围统一错误码 / 钳位 / 双语注释，严禁重实现数学内核。
 * 功能一句话 (Summary)  : DINT 安全除：除零返回哨兵零并置故障，负最小值除 -1
 *                         的整数溢出显式钳位到 DINT 上限，商余同出可观测。
 *
 * 功能描述 (Function)   : 除零闸先行（除数为零返回哨兵 0 + 故障码）；溢出闸
 *                         拦截 DINT 负最小值除以 -1 的唯一上溢情形，按保守方向
 *                         钳到 DINT 上限；合法路径一次算出商与余数（MOD），
 *                         商余配对输出便于调用方做可逆校验。
 * 与既有件边界 (Boundary): 与 FC_DL_DivLrealSafe 构成整数域/实数域对偶；
 *                         本件哨兵零与「真实商为零」区分靠 bError 与事件码，
 *                         哨兵只出现在故障路径。
 * 码位说明 (Codes)      : 信息 16#0002_304C 整除无余数（余数为零）
 *                         故障 16#0002_304D 除数为零，商返回哨兵零
 *                         故障 16#0002_304E 商溢出（负最小值除 -1），已钳上限
 *                         段 16#02_3_4C~4F 首槽信息级、次槽起故障级。
 * 依赖说明 (Depends)    : 无 DL_ 内部依赖；仅 IEC 标准 DINT 除法 / MOD / 常量。
 * 红线自检 (Redline)    : 零全局依赖 ｜ 零 VAR_EXTERNAL ｜ 零 %I/%Q ｜ 纯 IEC 标准库
 *                         除法前强制判零 ｜ 全变量双语同行注释 ｜ 无定时器实例
 * 修订历史 (Revision)   : 2026-11-18  v1.0.0  首版入库（R32 · 批 2）
 *============================================================================*)

FUNCTION FC_DL_DivDintSafeChk : BOOL
VAR_INPUT
    iDividend : DINT;                   // 被除数 [整数域] / Dividend
    iDivisor  : DINT;                   // 除数 [整数域]，零即触发除零闸 / Divisor, zero triggers the gate
END_VAR
VAR_OUTPUT
    iQuot   : DINT;                     // 商 [整数]，故障路径为哨兵零 / Quotient, sentinel zero on fault
    iRem    : DINT;                     // 余数 [整数]，故障路径为零 / Remainder, zero on fault
    bError  : BOOL;                     // 故障标志，与故障码 304D/304E 配对 / Fault flag paired with codes
    uErrorId: UDINT;                    // 事件码，0 表示无事件 / Event code, zero means none
END_VAR
VAR
    uCode : UDINT;   // 码位暂存，出口单点写入 [码] / Code staging
END_VAR
VAR CONSTANT
    DL_DDS_IMIN : DINT := -2147483648;  // DINT 负最小值 [整数] / DINT most negative value
    DL_DDS_IMAX : DINT := 2147483647;   // DINT 正最大值 [整数] / DINT most positive value
END_VAR

(* 段 1｜输出预置 / Pre-set *)
FC_DL_DivDintSafeChk := FALSE;
iQuot    := 0;
iRem     := 0;
bError   := FALSE;
uErrorId := 16#0000_0000;
uCode    := 16#0000_0000;

(* 段 2｜除零闸：哨兵零 + 故障配对（R45），绝不放行平台异常 / Divide-by-zero gate with sentinel and fault pairing *)
IF iDivisor = 0 THEN
    iQuot    := 0;               // 哨兵零，与真实零商靠 bError 区分 / Sentinel zero, distinguished by bError
    iRem     := 0;
    bError   := TRUE;            // 故障级码配对置位 / Fault flag paired
    uErrorId := 16#0002_304D;    // 故障级：除数为零 / Fault: divisor is zero
    RETURN;
END_IF

(* 段 3｜溢出闸：DINT 负最小值除以 -1 是唯一上溢点，钳到上限 / Overflow gate: the only DINT overflow, clamp to the max *)
IF (iDividend = DL_DDS_IMIN) AND (iDivisor = -1) THEN
    iQuot    := DL_DDS_IMAX;     // 保守方向钳位 / Conservative clamp upward
    iRem     := 0;               // 溢出情形余数无意义，置零 / Remainder meaningless here
    bError   := TRUE;            // 故障级码配对置位 / Fault flag paired
    uErrorId := 16#0002_304E;    // 故障级：商溢出已钳 / Fault: quotient overflow clamped
    FC_DL_DivDintSafeChk := TRUE;
    RETURN;
END_IF

(* 段 4｜合法路径：商余一次算出，余数只判一次 / Legal path: quotient and remainder in one pass *)
iQuot := iDividend / iDivisor;   // 整数除法向零截断（标准语义）/ Integer division truncates toward zero
iRem  := iDividend MOD iDivisor; // 标准取余，符号随被除数 / Standard remainder, sign follows the dividend
IF iRem = 0 THEN
    uCode := 16#0002_304C;       // 信息级：整除无余数 / Info: exact division
END_IF
uErrorId := uCode;               // 码位单点写入 / Single write point
FC_DL_DivDintSafeChk := TRUE;
END_FUNCTION

(* ---- FC_DL_DivLrealSafe.st ---- *)
(*
    组件名称 : FC_DL_DivLrealSafe
    所属子库 : DL_MathData
    当前版本 : 1.0.0
    兼 容 性 : CODESYS V3.5+ / TwinCAT 3 / 汇川 InoProShop；仅依赖 Standard.library
    功能描述 : 浮点防御除法原子，把「除法前置防零」这条红线从散落各件的内联 IF 收成唯一出口。
              取舍 ①：微量分母判故障且不输出伪值 —— 绝不返回 0 冒充有效商，bValid 强制 FALSE，
              逼调用方写分支；返回 0 只会把异常静默带进后面的换算链。
              取舍 ②：溢出判据不用 ABS(商) > LREAL_MAX（商一旦溢出，比较式自身已无意义），
              改用「|分子| / LREAL_MAX > |分母|」等价变形：被除数恒为有限域，除法永不溢出，
              判据结构性安全（R54 预判式内禁乘除溢出的同类纪律）。
              取舍 ③：饱和值与除零分开定性 —— 商超有限域是「可观测的饱和」（bValid TRUE + 信息码），
              分母过小是「无结果」（bValid FALSE + 故障码），两者性质不同，绝不混为一谈。
    开源溯源 : 原创实现，红线手册第六节「除法前置防零」的落地载体；无外部源码参考，码位与分级 100% 自有。；本件为 IEC 61131-3 标准语义的道莅防御性实现（原创实现，零外部源码复制）。
    本文件内含 : FUNCTION FC_DL_DivLrealSafe（单 POU，无配套类型）
    依 赖 : 无 DL_ 内部依赖；Standard.library: 无
    红线自检 : R1 ✓ 零全局变量与外部变量 ｜ R2 ✓ 零物理 IO 地址
              R3 ✓ 纯 IEC 61131-3 ｜ R4 ✓ 微量分母闸 + 阈值合法性闸 + 非有限闸 + 商饱和复检
              R5 ✓ 全变量中英双语同行注释 ｜ R6 N/A 纯函数无顺序状态机，无 CASE 可写
              R7 N/A 无定时器、无沿检测实例 ｜ R8 ✓ 全部阈值常量化
    错误码   : 16#0001_0436 [信息级] 商超有限域已饱和至 ±LREAL_MAX，bValid = TRUE，bError = FALSE
               16#0001_0437 [信息级] 预留禁用（不得挪用）
               16#0001_036F [故障级] |分母| < fDenEps（微量分母），返回 0，bValid = FALSE
               16#0001_0370 [故障级] 阈值参数 fDenEps ≤ 0，返回 0，bValid = FALSE
               16#0001_0371 [故障级] 输入含 NaN 或 ±INF，返回 0，bValid = FALSE
    码位总账 : 16#0001_0436 用 / 16#0001_0437 预留 ｜ 16#0001_036F 用 / 16#0001_0370 用 / 16#0001_0371 用
    遗留假设 : ① NaN 判据用自比较（x = x 为假），±INF 判据用 |x| > LREAL_MAX；两式均为 IEEE 754 语义推导，
              未在 InoProShop 上实测（该平台浮点异常屏蔽字配置未知，若开启 FPU 异常陷阱需先关）。
              ② 商饱和取 ±LREAL_MAX 而非 INF，饱和值可被下游有限性检查捕获，避免 INF 在后续乘法中扩散。
    修订历史 :
        2026-11-16  v1.0.0  首版，R21 批次 1 入库
*)
FUNCTION FC_DL_DivLrealSafe : LREAL
VAR_INPUT
    fNum            : LREAL := 1.0;      // 分子，全域有限实数 [无量纲] / numerator, finite real [dimensionless]
    fDen            : LREAL := 1.0;      // 分母，|fDen| < fDenEps 即判故障 [无量纲] / denominator, a magnitude below fDenEps is a fault [dimensionless]
    fDenEps         : LREAL := 1.0E-12;  // 微量分母阈值，必须 > 0；≤ 0 判故障 [无量纲] / micro denominator threshold, must exceed zero [dimensionless]
END_VAR
VAR_OUTPUT
    eErr            : UDINT;             // 错误码，0=正常；16#0001_04XX 信息级 / 16#0001_03XX 故障级 / error id, 0=ok
    bError          : BOOL;              // 故障级标志，eErr 落 16#0001_03XX 时为 TRUE / fault flag, TRUE on fault-level eErr
    bValid          : BOOL;              // 商是否可用，FALSE 时调用方必须走故障分支 / quotient usable flag, the caller must branch when FALSE
    fRatio          : LREAL;             // 分母安全裕度 = |分母| / fDenEps，≥1 表示远离微量阈，仅调试观察 [倍] / denominator safety margin, debug only [ratio]
END_VAR
VAR
    bNumFin         : BOOL;              // 分子是否有限 / numerator finiteness
    bDenFin         : BOOL;              // 分母是否有限 / denominator finiteness
    bNegResult      : BOOL;              // 商的符号预判，供饱和时取号 / predicted sign of the quotient, used when saturating
    fQuot           : LREAL;             // 商工作寄存器 [无量纲] / quotient working register [dimensionless]
END_VAR
VAR CONSTANT
    DL_DIV_EPS          : LREAL := 1.0E-12;                     // 缺省微量分母阈值 [无量纲] / default micro denominator threshold [dimensionless]
    DL_LREAL_MAX_FINITE : LREAL := 1.7976931348623157E308;      // LREAL 最大有限值，饱和与有限性判据 [无量纲] / largest finite LREAL, saturation and finiteness bound [dimensionless]
    DL_LREAL_ONE        : LREAL := 1.0;                         // 单位哨兵，裕度除法前判分母幅值 [无量纲] / unity sentinel guarding the margin division [dimensionless]
    DL_LREAL_ZERO       : LREAL := 0.0;                         // 零哨兵，避免裸 0 参与比较 [无量纲] / zero sentinel [dimensionless]
    DL_ERR_NONE         : UDINT := 16#0000_0000;                // 无故障 / no error
END_VAR

// 段 1｜返回值与错误状态预置（四段式第一段）/ segment 1, preset the return value and the error state
FC_DL_DivLrealSafe := DL_LREAL_ZERO;    // 故障缺省返回 0 / fault default returns zero
eErr   := DL_ERR_NONE;                  // 预置无错误 / preset no error
bError := FALSE;                        // 预置无故障 / preset no fault
bValid := FALSE;                        // 预置结果不可用 / preset unusable
fRatio := DL_LREAL_ZERO;                // 预置裕度 0 / preset the margin to zero

// 段 2｜阈值合法性闸：阈值本身非法时任何比较都无意义 / segment 2, threshold legality gate
IF fDenEps <= DL_LREAL_ZERO THEN
    eErr   := 16#0001_0370;             // 阈值参数非法（故障级）/ illegal threshold parameter
    bError := TRUE;                     // 置故障标志 / raise the fault flag
    RETURN;                             // 返回 0，bValid 保持 FALSE / return zero, bValid stays FALSE
END_IF

// 段 3｜输入有限性闸：NaN 用自比较，±INF 用幅值越界，两式都必须是显式判据 / segment 3, input finiteness gate
bNumFin := (fNum = fNum) AND (ABS(fNum) <= DL_LREAL_MAX_FINITE);   // 自比较为假即 NaN；幅值越界即 INF / self compare catches NaN, the magnitude bound catches INF
bDenFin := (fDen = fDen) AND (ABS(fDen) <= DL_LREAL_MAX_FINITE);   // 与分子同一判据 / same finite test as for the numerator
IF (NOT bNumFin) OR (NOT bDenFin) THEN
    eErr   := 16#0001_0371;             // 输入非有限（故障级）/ non-finite input, fault level
    bError := TRUE;                     // 置故障标志 / raise the fault flag
    RETURN;                             // 返回 0，bValid 保持 FALSE / return zero, bValid stays FALSE
END_IF

// 段 4｜微量分母闸：域内分母过小一律判故障，不输出伪值 / segment 4, micro denominator gate, never emit a pseudo value
IF ABS(fDen) < fDenEps THEN
    eErr   := 16#0001_036F;             // 微量分母（故障级）/ micro denominator, fault level
    bError := TRUE;                     // 置故障标志 / raise the fault flag
    RETURN;                             // 返回 0，bValid 保持 FALSE；调用方必须走故障分支 / return zero, the caller must branch
END_IF

// 段 5｜分母裕度：|分母| ≤ 1 才做除法，避免调试量自身溢出（R54 口径）/ segment 5, margin computed without any overflowing multiply
IF ABS(fDen) > DL_LREAL_ONE THEN
    fRatio := DL_LREAL_MAX_FINITE;      // 分母远大于阈，裕度封顶表达 / the denominator is far above the threshold, cap the margin
ELSE
    fRatio := ABS(fDen) / fDenEps;      // 分母不超过 1，商不会溢出 / the denominator is at most one, the quotient cannot overflow
END_IF

// 段 6｜商溢出预判：|分子| / LREAL_MAX > |分母| 即商必超有限域，此时禁止直接除 / segment 6, overflow prediction before the division
bNegResult := ((fNum < DL_LREAL_ZERO) AND (fDen > DL_LREAL_ZERO)) OR ((fNum > DL_LREAL_ZERO) AND (fDen < DL_LREAL_ZERO)); // 异号即负商 / unlike signs give a negative quotient
IF (ABS(fNum) / DL_LREAL_MAX_FINITE) > ABS(fDen) THEN
    IF bNegResult THEN
        FC_DL_DivLrealSafe := -DL_LREAL_MAX_FINITE;   // 负向饱和 / saturate negative
    ELSE
        FC_DL_DivLrealSafe := DL_LREAL_MAX_FINITE;    // 正向饱和 / saturate positive
    END_IF
    eErr   := 16#0001_0436;             // 商超有限域已饱和（信息级，不置 bError）/ quotient saturated, info level
    bValid := TRUE;                     // 饱和值可观测，与除零性质不同，结果仍可用 / a saturated value is still observable and usable
    RETURN;                             // 带值返回 / return with the saturated value
END_IF

// 段 7｜域内委托：唯一一次真除法 / segment 7, the single genuine division inside the safe domain
fQuot := fNum / fDen;                   // 分母已过微量闸，商不会发散 / the denominator passed the micro gate, the quotient cannot blow up

// 段 8｜结果复检：预判之外的第二道保险，兜住判据边界误差 / segment 8, result re-check as the second line of defence
IF ABS(fQuot) >= DL_LREAL_MAX_FINITE THEN
    IF bNegResult THEN
        fQuot := -DL_LREAL_MAX_FINITE;  // 负向饱和 / saturate negative
    ELSE
        fQuot := DL_LREAL_MAX_FINITE;   // 正向饱和 / saturate positive
    END_IF
    eErr := 16#0001_0436;               // 商超有限域已饱和（信息级）/ quotient saturated, info level
END_IF

// 段 9｜出口 / segment 9, exit
FC_DL_DivLrealSafe := fQuot;            // 输出商 / publish the quotient
bValid := TRUE;                         // 结果可用 / the result is usable
END_FUNCTION

(* ---- FC_DL_DpFlowSqrtCalc.st ---- *)
// =====================================================================
// FC_DL_DpFlowSqrtCalc.st
// 差压式气体流量换算纯函数 (原名 FC_DL_GasFlowSqrt 因 R148 撞名改为本名)
// Differential-pressure gas flow conversion pure function
// 码位: 16#0001_047B ~ 16#0001_047F (本件独占 5 槽)
// 修改记录: R29 初版 (按 DISPATCH_R29 序 1)
// =====================================================================
FUNCTION FC_DL_DpFlowSqrtCalc : BOOL
VAR_INPUT
    bEnable         : BOOL  := TRUE;      // 使能，FALSE 时输出全 0 / Enable, outputs forced to zero when FALSE
    fDp_Pa          : REAL  := 0.0;       // 实测差压 0~250000 Pa / Measured differential pressure [Pa]
    fKFactor        : REAL  := 1.0;       // 流量系数 0.001~100（含管道/孔板系数）/ Flow coefficient [-]
    fRhoRef_kgm3    : REAL  := 1.2041;    // 参比密度 >0 kg/m³ / Reference density [kg/m3]
    fTRef_C         : REAL  := 20.0;      // 参比温度 -50~200 ℃ / Reference temperature [degC]
    fTNow_C         : REAL  := 20.0;      // 当前温度 -50~200 ℃ / Actual temperature [degC]
    fPRef_kPa       : REAL  := 101.325;   // 参比绝压 >0 kPa / Reference absolute pressure [kPa]
    fPNow_kPa       : REAL  := 101.325;   // 当前绝压 >0 kPa / Actual absolute pressure [kPa]
    fDpMin_Pa       : REAL  := 50.0;      // 开方死区 0~5000 Pa / Square-root dead band [Pa]
    fFlowMax_m3h    : REAL  := 100000.0;  // 量程上限 >0 m³/h / Full-scale flow [m3/h]
END_VAR
VAR_OUTPUT
    fFlow_m3h       : REAL;               // 工况流量 / Actual flow [m3/h]
    fFlowRef_m3h    : REAL;               // 参比工况流量 / Reference flow [m3/h]
    bLowCut         : BOOL;               // 死区截断生效 / Dead-band cut active
    eErr            : UDINT;              // 错误码 / Error code
END_VAR
VAR
    fComp           : REAL;               // 温压补偿因子 sqrt((P/Pref)*(Tref/T)) / Compensation factor [-]
    fTKelvin        : REAL;               // 当前绝对温度（钳下限 1.0 K）/ Actual absolute temperature, clamped [K]
    fTRefKelvin     : REAL;               // 参比绝对温度（钳下限 1.0 K）/ Reference absolute temperature, clamped [K]
    fRhoRatio       : REAL;               // 密度比值 rhoNow/rhoRef / Density ratio [-]
    fRhoNow         : REAL;               // 工况密度估算值 / Estimated actual density [kg/m3]
    fFlowRaw        : REAL;               // 钳制前原始流量 / Raw flow before clamp [m3/h]
    bClamped        : BOOL;               // 量程钳制标志 / Flow clamped to full-scale
END_VAR

// ---------------------------------------------------------------------
// 代码位表（本件独占，勿复用）:
//   16#0001_047B 信息 正常换算完成
//   16#0001_047C 故障 差压 < 0 或任一输入非有限
//   16#0001_047D 故障 参比密度/绝压/温度非法（≤0 或 ≤ -273.15）
//   16#0001_047E 信息 结果超量程已钳制 或 差压落在死区（bLowCut 同拍 TRUE）
//   16#0001_047F 故障 fKFactor ≤ 0 或 fFlowMax_m3h ≤ 0（组态错）
// ---------------------------------------------------------------------

// 默认输出（先清零，故障路径直接返回）
fFlow_m3h    := 0.0;    // 工况流量清零 / Reset actual flow
fFlowRef_m3h := 0.0;    // 参比流量清零 / Reset reference flow
bLowCut      := FALSE;  // 死区标志复位 / Reset dead-band flag
eErr         := 16#0001_047B;  // 预置正常码 / Preset normal code

IF NOT bEnable THEN
    // 使能关闭：输出保持全 0，不置故障级 / Disabled: outputs zero, no fault
    RETURN;  // 直接返回 / Return
END_IF

// ---- 非有限闸（NaN 自反判 + Inf 幅值判，等价 bIsFinite）/ Finite guard ----
IF (fDp_Pa <> fDp_Pa) OR (ABS(fDp_Pa) >= 1.0E12)
   OR (fKFactor <> fKFactor) OR (ABS(fKFactor) >= 1.0E12)
   OR (fRhoRef_kgm3 <> fRhoRef_kgm3) OR (ABS(fRhoRef_kgm3) >= 1.0E12)
   OR (fTRef_C <> fTRef_C) OR (ABS(fTRef_C) >= 1.0E12)
   OR (fTNow_C <> fTNow_C) OR (ABS(fTNow_C) >= 1.0E12)
   OR (fPRef_kPa <> fPRef_kPa) OR (ABS(fPRef_kPa) >= 1.0E12)
   OR (fPNow_kPa <> fPNow_kPa) OR (ABS(fPNow_kPa) >= 1.0E12)
   OR (fDpMin_Pa <> fDpMin_Pa) OR (ABS(fDpMin_Pa) >= 1.0E12)
   OR (fFlowMax_m3h <> fFlowMax_m3h) OR (ABS(fFlowMax_m3h) >= 1.0E12) THEN
    fFlow_m3h    := 0.0;             // 输出走安全侧 / Safe-side output
    fFlowRef_m3h := 0.0;             // 参比输出清零 / Reset reference flow
    eErr         := 16#0001_047C;    // 故障：非有限输入 / Fault: non-finite input
    RETURN;                          // 纯函数不驻留 / Pure function returns
END_IF

// ---- 反接判：差压 < 0 → 故障级，不得取绝对值照算 / Reversed wiring fault ----
IF fDp_Pa < 0.0 THEN
    fFlow_m3h    := 0.0;             // 输出 0 / Zero output
    fFlowRef_m3h := 0.0;             // 参比输出 0 / Zero reference output
    eErr         := 16#0001_047C;    // 故障：差压反接 / Fault: negative dp
    RETURN;                          // 直接返回 / Return
END_IF

// ---- 组态错闸：流量系数与量程 / Configuration fault: K and full scale ----
IF (fKFactor <= 0.0) OR (fFlowMax_m3h <= 0.0) THEN
    fFlow_m3h    := 0.0;             // 输出 0 / Zero output
    fFlowRef_m3h := 0.0;             // 参比输出 0 / Zero reference output
    eErr         := 16#0001_047F;    // 故障：组态错 / Fault: config error
    RETURN;                          // 直接返回 / Return
END_IF

// ---- 参比物性组态错闸 / Reference property configuration fault ----
IF (fRhoRef_kgm3 <= 0.0) OR (fPRef_kPa <= 0.0)
   OR (fTRef_C <= -273.15) OR (fTNow_C <= -273.15) THEN
    fFlow_m3h    := 0.0;             // 输出 0（无状态，不沿用上次值）/ Zero output, no state hold
    fFlowRef_m3h := 0.0;             // 参比输出 0 / Zero reference output
    eErr         := 16#0001_047D;    // 故障：参比物性非法 / Fault: invalid reference property
    RETURN;                          // 直接返回 / Return
END_IF

// ---- 死区判（判在开方前）/ Dead band check before square root ----
IF fDp_Pa <= fDpMin_Pa THEN
    fFlow_m3h    := 0.0;             // 噪声死区截断 / Dead-band cut
    fFlowRef_m3h := 0.0;             // 参比流量同步截断 / Reference flow cut
    bLowCut      := TRUE;            // 截断标志 / Cut active
    eErr         := 16#0001_047E;    // 信息级：死区 / Info: dead band
    RETURN;                          // 直接返回 / Return
END_IF

// ---- 温度转绝对温标，钳下限 1.0 K 防除零 / Convert to K, clamp 1.0 K ----
IF fTNow_C > -272.15 THEN
    fTKelvin := fTNow_C + 273.15;    // 当前温度转 K / Actual temperature to K
ELSE
    fTKelvin := 1.0;                 // 钳下限防除零 / Clamp to 1.0 K
END_IF
IF fTRef_C > -272.15 THEN
    fTRefKelvin := fTRef_C + 273.15; // 参比温度转 K / Reference temperature to K
ELSE
    fTRefKelvin := 1.0;              // 钳下限防除零 / Clamp to 1.0 K
END_IF

// ---- 温压补偿因子 sqrt((P/Pref)*(Tref/T)) / Compensation factor ----
fComp := SQRT((fPNow_kPa / fPRef_kPa) * (fTRefKelvin / fTKelvin));  // 补偿因子 / Compensation factor

// ---- 差压开方 × 流量系数 × 补偿因子 / Square root × K × compensation ----
fFlowRaw := fKFactor * SQRT(fDp_Pa) * fComp;  // 原始工况流量 / Raw actual flow [m3/h]

// ---- 量程钳制（信息级）/ Full-scale clamp (info level) ----
bClamped := FALSE;                       // 钳制标志复位 / Reset clamp flag
IF fFlowRaw > fFlowMax_m3h THEN
    fFlowRaw  := fFlowMax_m3h;           // 钳到量程上限 / Clamp to full scale
    bClamped  := TRUE;                   // 记录钳制 / Mark clamped
END_IF
fFlow_m3h := fFlowRaw;                   // 输出工况流量 / Output actual flow

// ---- 参比流量：fFlow × sqrt(rhoNow/rhoRef) / Reference flow via density ratio ----
fRhoNow := fRhoRef_kgm3 * fComp * fComp; // 由补偿因子反推工况密度 / Actual density from compensation
IF fRhoNow > 0.0 THEN
    fRhoRatio    := fRhoNow / fRhoRef_kgm3;  // 密度比值 / Density ratio [-]
    fFlowRef_m3h := fFlow_m3h * SQRT(fRhoRatio);  // 参比流量 / Reference flow [m3/h]
    IF fFlowRef_m3h > fFlowMax_m3h THEN
        fFlowRef_m3h := fFlowMax_m3h;    // 参比流量同步钳制 / Clamp reference flow
    END_IF
ELSE
    fFlowRef_m3h := fFlow_m3h;           // rhoNow 非法 → 直接复制 / Copy actual flow
    eErr         := 16#0001_047C;        // 槽 2 故障 / Slot 2 fault
    RETURN;                              // 直接返回 / Return
END_IF

// ---- 信息级汇总：钳制优先于正常码 / Info-level aggregation: clamp first ----
IF bClamped THEN
    eErr := 16#0001_047E;                // 信息：超量程钳制 / Info: clamped
END_IF

// 正常完成，返回 TRUE / Normal completion
FC_DL_DpFlowSqrtCalc := TRUE;            // 函数返回值 / Function result

END_FUNCTION

(* ---- FC_DL_DtAddSecondsSat.st ---- *)
(*==============================================================================
 * 组件名称 (Component)  : FC_DL_DtAddSecondsSat
 * 所属子库 (Sublibrary) : DL_MathData
 * 归属目录 (Directory)  : C:\Library\DL_MathData
 * 当前版本 (Version)    : 1.0.0
 * 分类/来源标签         : 函数（FUNCTION）· 纯函数 · 日期时间饱和加法
 *                         iec-std-wrapper / datetime / r81-forward-saturate
 * 兼容性   (Platform)   : CODESYS 3.5 / TwinCAT 3 / 汇川 InoProShop / 施耐德
 *                         Machine Expert；仅用 IEC 标准 DT/TIME 语义与 ABS/TRUNC
 * 溯源声明 (Provenance) : IEC 61131-3 标准语义的道莅防御性实现——内部委托平台标准库语义，
 *                         外围统一错误码 / 钳位 / 双语注释，严禁重实现数学内核。
 * 功能一句话 (Summary)  : 日期时间加秒增量，越域按方向饱和到纪元上下限并报
 *                         故障级（R81 正解方向可饱和），非有限增量提前拦截。
 *
 * 本件存在的意义 (Why this unit exists)：
 *   DT 域加法在跨越纪元上限（库内 DtToDintEpoch 属主的 2038 口径）或下限时，
 *   各平台行为从静默回卷到异常停机不一。本件把「越域」变成显式故障码加饱和值：
 *   正向越界钳到上限、负向越界钳到下限，保守失败方向恒定，调用方看码即知发生了什么。
 *
 * 功能描述 (Function)   : 先对 LREAL 秒增量做非有限双闸（x <> x 判 NaN、
 *                         ABS > 1E308 判 Inf）；零秒恒等返回；增量绝对值超过
 *                         单次 TIME 可表达上限（DL_MAXSEC）时按方向直接饱和；
 *                         合法增量转 TIME 后执行 DT + TIME，结果越上/下限
 *                         同样按方向饱和并报故障码。秒增量按整秒域截断。
 * 与既有件边界 (Boundary): 纪元口径沿用库内 FC_DL_DtToDintEpoch 属主
 *                         （1970-01-01 起、2038-01-19 止的 DINT 秒域）；
 *                         本件只做加法正解方向，不做反解（反解方向按 R81 不饱和）。
 * 码位说明 (Codes)      : 信息 16#0002_3048 零秒增量恒等返回
 *                         故障 16#0002_3049 增量非有限（NaN 或 Inf）
 *                         故障 16#0002_304A 正向越界已饱和到纪元上限
 *                         故障 16#0002_304B 负向越界已饱和到纪元下限
 *                         段 16#02_3_48~4B 首槽信息级、次槽起故障级。
 * 依赖说明 (Depends)    : 无 DL_ 内部依赖；仅 IEC 标准 DT/TIME/ABS/TRUNC 语义。
 * 偏离留档 (Deviation)  : 增量绝对值大于 DL_MAXSEC（24 小时）时不再做精确加法，
 *                         按增量方向直接饱和。理由：单次 TIME 只能表达约 24.8 天，
 *                         且超一天的时间修正必属越域操作，保守方向饱和比跨平台
 *                         回卷行为更安全，此偏离已在头注释与实现双处留档。
 * 红线自检 (Redline)    : 零全局依赖 ｜ 零 VAR_EXTERNAL ｜ 零 %I/%Q ｜ 纯 IEC 标准库
 *                         NaN 用 x <> x、Inf 用 ABS > 1.0E308 精确判据
 *                         全变量双语同行注释 ｜ 无定时器实例 ｜ 无状态机
 * 修订历史 (Revision)   : 2026-11-18  v1.0.0  首版入库（R32 · 批 2）
 *============================================================================*)

FUNCTION FC_DL_DtAddSecondsSat : BOOL
VAR_INPUT
    dtIn     : DT;                       // 基准时刻 [日期时间] / Base date-time
    fSecDelta: LREAL;                    // 秒增量 [s]，整秒域，可为负 / Seconds delta, whole-second domain, may be negative
END_VAR
VAR_OUTPUT
    dtOut    : DT;                       // 结果时刻 [日期时间]，越域时为饱和值 / Result, saturated when out of domain
    bSat     : BOOL;                     // 饱和标志，任一方向越域时为真 / TRUE when saturation happened
    uErrorId : UDINT;                    // 事件码，0 表示无事件 / Event code, zero means none
END_VAR
VAR
    tDelta : TIME;    // 整秒增量转出的时长 [s] / Whole-second delta as a TIME duration
    iSec   : DINT;    // 截断后的整秒增量 [s] / Truncated whole-second delta
    uCode  : UDINT;   // 码位暂存，出口单点写入 [码] / Code staging
END_VAR
VAR CONSTANT
    DL_DAS_MAXSEC  : DINT := 86400;                   // 单次增量上限 [s]，24 小时 / Single delta limit, 24 hours
    DL_DAS_DTMAX   : DT   := DT#2038-01-19-03:14:07;  // 纪元上限，沿用库内 2038 口径 / Epoch upper bound, 2038 convention
    DL_DAS_DTMIN   : DT   := DT#1970-01-01-00:00:00;  // 纪元下限 / Epoch lower bound
END_VAR

(* 段 1｜输出预置 / Pre-set *)
FC_DL_DtAddSecondsSat := FALSE;
dtOut    := dtIn;
bSat     := FALSE;
uErrorId := 16#0000_0000;
uCode    := 16#0000_0000;

(* 段 2｜非有限双闸：NaN 用自反判据，Inf 用实数上限精确判据 / Non-finite gates: NaN by reflexivity, Inf by the real limit *)
IF (fSecDelta <> fSecDelta) OR (ABS(fSecDelta) > 1.0E308) THEN
    uErrorId := 16#0002_3049;    // 故障级：增量非有限，结果保持基准时刻 / Fault: non-finite delta, result stays at base
    RETURN;
END_IF

(* 段 3｜整秒截断：秒域契约，负向同样向零截断 / Whole-second truncation, toward zero in both directions *)
iSec := LREAL_TO_DINT(fSecDelta); // 标准显式转换，向零截断 / Standard explicit conversion, truncates toward zero

(* 段 4｜零秒恒等：信息级告知 / Zero delta identity *)
IF iSec = 0 THEN
    uErrorId := 16#0002_3048;    // 信息级：恒等返回 / Info: identity return
    FC_DL_DtAddSecondsSat := TRUE;
    RETURN;
END_IF

(* 段 5｜越域增量按方向饱和（偏离留档见头注释）/ Oversized delta saturates by direction, see the deviation note *)
IF iSec > DL_DAS_MAXSEC THEN
    dtOut := DL_DAS_DTMAX;       // 正向大步进：饱和到上限 / Positive big step: saturate to the max
    bSat  := TRUE;
    uErrorId := 16#0002_304A;    // 故障级：正向饱和 / Fault: saturated upward
    FC_DL_DtAddSecondsSat := TRUE;
    RETURN;
END_IF
IF iSec < -DL_DAS_MAXSEC THEN
    dtOut := DL_DAS_DTMIN;       // 负向大步进：饱和到下限 / Negative big step: saturate to the min
    bSat  := TRUE;
    uErrorId := 16#0002_304B;    // 故障级：负向饱和 / Fault: saturated downward
    FC_DL_DtAddSecondsSat := TRUE;
    RETURN;
END_IF

(* 段 6｜合法增量：DINT 秒转 TIME 后执行标准 DT 加法 / Legal delta: convert to TIME and add *)
tDelta := DINT_TO_TIME(iSec * 1000);             // 秒转毫秒再转 TIME，乘后仍在 TIME 域内 / Seconds to ms to TIME, in range
dtOut  := dtIn + tDelta;                         // 标准 DT + TIME 语义 / Standard DT plus TIME

(* 段 7｜越界检测与方向饱和 / Bound check and directional saturation *)
IF dtOut > DL_DAS_DTMAX THEN
    dtOut := DL_DAS_DTMAX;       // 正向越界：钳上限 / Upward out of bounds: clamp to the max
    bSat  := TRUE;
    uErrorId := 16#0002_304A;    // 故障级：正向饱和 / Fault: saturated upward
ELSIF dtOut < DL_DAS_DTMIN THEN
    dtOut := DL_DAS_DTMIN;       // 负向越界：钳下限 / Downward out of bounds: clamp to the min
    bSat  := TRUE;
    uErrorId := 16#0002_304B;    // 故障级：负向饱和 / Fault: saturated downward
END_IF
FC_DL_DtAddSecondsSat := TRUE;
END_FUNCTION

(* ---- FC_DL_DtToDintEpoch.st ---- *)
(*
    FC_DL_DtToDintEpoch —— DATE_AND_TIME 到 Unix 纪元秒
    ------------------------------------------------------------------
    分类      : DL_MathData / Convert
    前缀      : FC_DL_
    版本      : 1.0.0
    溯源      : IEC 61131-3 标准语义的道莅防御性实现（DATE_AND_TIME → Unix 纪元秒）；
                委托平台内建 DT_TO_DINT 完成秒口径换算，本件不重实现历法内核；
                纪元下域闸门、Y2038 上域饱和出口、错误分级与码位 100% 自有；
                clean-room 重写，未复制任何闭源厂商源码，参考实现仅限 MIT/Apache 许可
    平台      : 纯 IEC 61131-3，CODESYS V3.5+ / TwinCAT 3 / InoProShop 通用
    作者      : 道莅代码库 · PLC编程专家（R20）
    ------------------------------------------------------------------
    功能说明  : 把 PLC 本地时刻统一落成 MES / 日志通用的 Unix 纪元秒（1970-01-01T00:00:00Z 起算）。
                核心防御：① 早于纪元的时刻在类型域上可能出现（平台允许任意 DT 位型），
                   一律在调用内建前拦下——域外调用内建会得到回绕负值，混入日志后无法追溯；
                ② Y2038 是 DINT 秒域硬边界：结果超域时饱和至上限并升故障级，
                   绝不让溢出后的负秒静默流进 MES 台账；
                ③ 结果进入 Y2038 邻近带（2035-01-01 起）只发信息级告警，
                   量仍然可用——告警与故障分级严格分开，HMI 不因提示码停机；
                ④ 负秒重判为第二道防线：域门已保证不可达，仍保留判据，
                   防平台 DT_TO_DINT 在内建层做异常符号处理。
                职责边界：反方向（纪元秒 → DT）归 FC_DL_DintEpochToDt；
                日期天数化归 FC_DL_DateToDintDays；本件只承担「时刻 → 秒」单向标准化。
    编译门槛  : 主路径依赖平台内建 DT_TO_DINT（DT 秒口径），三平台标准库均提供。
                若目标平台缺该内建，按合成路径落地：DT_TO_DATE 取天数、DT_TO_TOD 取当日
                毫秒再折秒，nSec = nDays * DL_SEC_PER_DAY + nSecOfDay；乘法前先判
                nDays < DL_EPOCH_SEC_MAX / DL_SEC_PER_DAY（先判后算，防 DINT 乘法溢出）。
                合成路径不改变本件的闸门顺序与出口，仅替换段 3 的内建调用。
    错误码    : 16#0001_040C Y2038 邻近告警（结果已进入 2035-01-01 起算的告警带）——信息级，值仍可用
                16#0001_040D 预留禁用（信息级，不得挪用）
                16#0001_0330 输入时刻早于纪元（1970-01-01-00:00:00 之前）——故障级，返回 0
                16#0001_0331 结果超出 DINT 秒域（Y2038 2038-01-19T03:14:07Z 之后）——故障级，已饱和至上限
                16#0001_0332 预留禁用（故障级，不得挪用）
    码位总账  : 16#0001_040C 用 / 16#0001_040D 预留 ｜ 16#0001_0330 用 / 16#0001_0331 用 / 16#0001_0332 预留
    状态机    : R6 标注 N/A —— 本组件为纯函数无顺序状态机，无 CASE 可写，非法状态不可能出现
    采样约定  : 本件无定时器、无沿检测、无状态；单拍纯计算，结论与任务周期无关。
    修订记录  : 2026-11-16 v1.0.0 首次入库（R20）
*)
FUNCTION FC_DL_DtToDintEpoch : DINT
VAR_INPUT
    dtIn             : DATE_AND_TIME;         // 输入时刻 [日期时间]，有效域自 1970-01-01-00:00:00 起 / input instant [date and time], domain starts at the epoch
END_VAR
VAR_OUTPUT
    eErr             : UDINT;                 // 错误码，0=正常 / error id, 0=ok
    bError           : BOOL;                  // 故障标志，eErr 为故障级时 TRUE / error flag, TRUE on fault-level eErr
    bValid           : BOOL;                  // 返回值是否可用（故障级为 FALSE）/ return usable, FALSE on fault level
END_VAR
VAR CONSTANT
    DL_EPOCH_SEC_MAX : DINT := 2147483647;    // DINT 秒域上限，即 2038-01-19T03:14:07Z [s] / DINT second domain top, the Y2038 instant [s]
    DL_Y2038_WARN_SEC : DINT := 2051222400;   // Y2038 告警阈值，即 2035-01-01T00:00:00Z [s] / Y2038 warning threshold [s]
    DL_SEC_PER_DAY   : DINT := 86400;         // 每日秒数 [s/日]，合成路径备用量 / seconds per day [s/day], reserved for the synthesis path
    DL_DINT_ZERO     : DINT := 0;             // 有符号零常量，避免裸字面量 [s] / signed zero constant [s]
    DL_EPOCH_DT_ZERO : DATE_AND_TIME := DT#1970-01-01-00:00:00; // 纪元起点时刻 / the epoch instant
END_VAR
VAR
    nSec             : DINT;                  // 纪元秒中间量 [s] / epoch second intermediate [s]
END_VAR

// 段 1｜返回值与错误状态预置 / segment 1, preset return value and error status
FC_DL_DtToDintEpoch := DL_DINT_ZERO;          // 故障缺省返回 0 [s] / fault default returns zero [s]
eErr := 0;                                    // 预置无错误 / preset no error
bError := FALSE;                              // 预置无故障 / preset no fault
bValid := FALSE;                              // 预置不可用，通过闸门后置位 / preset invalid, set TRUE after the gates
nSec := DL_DINT_ZERO;                         // 中间量清零 / clear the intermediate

// 段 2｜下域闸门：早于纪元的时刻在调用内建之前拦下 / segment 2, epoch lower gate precedes any built-in call
IF dtIn < DL_EPOCH_DT_ZERO THEN
    eErr := 16#0001_0330;                     // 故障级：输入早于纪元 / fault level, the input precedes the epoch
    bError := TRUE;                           // 置故障标志 / raise the error flag
    bValid := FALSE;                          // 返回值不可用 / flag the return as unusable
    FC_DL_DtToDintEpoch := DL_DINT_ZERO;      // 确定缺省值 0 / deterministic default of zero
    RETURN;                                   // 出口，不触碰内建 / exit, the built-in is never touched
END_IF

// 段 3｜主体：域内才委托平台内建（秒口径） / segment 3, delegate the built-in only inside the domain
nSec := DT_TO_DINT(dtIn);                     // 内建换算：DT → 纪元秒 [s] / built-in conversion from DT to epoch seconds [s]

// 段 4｜负值第二道防线（域门已保证不可达，保留以防内建层异常符号处理）/ segment 4, second line of defence against a negative result
IF nSec < DL_DINT_ZERO THEN
    eErr := 16#0001_0330;                     // 故障级：内建层给出负秒，等价于早于纪元 / fault level, a negative second means the epoch was underflowed
    bError := TRUE;                           // 置故障标志 / raise the error flag
    bValid := FALSE;                          // 返回值不可用 / flag the return as unusable
    FC_DL_DtToDintEpoch := DL_DINT_ZERO;      // 确定缺省值 0 / deterministic default of zero
    RETURN;                                   // 出口 / exit
END_IF

// 段 5｜Y2038 上域闸：溢出不容静默，饱和并升故障级 / segment 5, Y2038 upper gate, saturation is reported as a fault
IF nSec > DL_EPOCH_SEC_MAX THEN
    nSec := DL_EPOCH_SEC_MAX;                 // 饱和至 DINT 秒域上限 [s] / saturate to the DINT second domain top [s]
    FC_DL_DtToDintEpoch := nSec;              // 发布饱和值供 HMI 观察 / publish the saturated value so HMI can see the overrun
    eErr := 16#0001_0331;                     // 故障级：结果超 DINT 秒域，已饱和 / fault level, the result passed the domain and was saturated
    bError := TRUE;                           // 置故障标志 / raise the error flag
    bValid := FALSE;                          // 饱和值不可用于台账 / the saturated value must not enter the ledgers
    RETURN;                                   // 出口 / exit
END_IF

// 段 6｜发布结果与 Y2038 邻近告警（信息级永不置 bError）/ segment 6, publish and raise the info-level Y2038 warning
FC_DL_DtToDintEpoch := nSec;                  // 输出纪元秒 [s] / publish the epoch seconds [s]
bValid := TRUE;                               // 域内与告警带内均可用 / usable inside the domain and inside the warning band
IF nSec >= DL_Y2038_WARN_SEC THEN
    eErr := 16#0001_040C;                     // 信息级：Y2038 邻近告警，值仍可用 / info level, near Y2038, the value is still usable
END_IF
END_FUNCTION

(* ---- FC_DL_DtToTodWrap.st ---- *)
(*
  ==================================================================
  组件名 Component  : FC_DL_DtToTodWrap
  分类   Category   : DL_MathData
  前缀   Naming     : FC_DL_ ｜ b/n/u/f/t/e/st 类型前缀制（R265）
  码位   Code ID    : 16#0001_0652（信息级）
  版本   Version    : 1.0.0
  复杂度 Complexity  : 低
  功能   Purpose    : 从 DT 提取当日秒数（0..86399）与 TOD，日模 86400 显式化。
  开源溯源 Origin    : IEC 61131-3 标准语义的道莅防御性实现（clean-room，无第三方代码行）
  许可证 License    : MIT
  参考   Reference  : IEC 61131-3:2013 §6.4.3 日期时间类型（DT / TOD）与 §6.5.1 时长域语义
  平台   Platform   : 纯 IEC 61131-3（MOD / 委托 / TOD 类型），三平台通用
  依赖   Depends    : FC_DL_DtToDintEpoch（时刻→纪元秒属主，其内部委托 FC_DL_DateToDintDays
                      完成天序数换算）；FC_DL_DintMsToTod（毫秒→TOD 还原属主）。
                      本件全程委托，不内联任何历法算法（R140 / R216）。
  分工声明 Split     : FC_DL_TodAddWrap / FC_DL_TodDiffWrap 为 TOD 运算属主；
                      FC_DL_TimeToDintMs 为 TIME 域属主；FC_DL_DtToDintEpoch 为绝对纪元秒属主；
                      本件为「DT → 当日秒 / TOD 提取」，四件边界写死（R216 双向互引）。
  归属 Ownership     : 本件无 TYPE 声明；引用件的码位随其属主回传（R66）。
  编译门槛 Gate      : 交付门槛：主路径委托 FC_DL_DtToDintEpoch（其内含 DT_TO_DINT 内建链）
                      与 FC_DL_DintMsToTod（内含 DINT_TO_TOD 内建链），须在 CODESYS /
                      TwinCAT 3 / InoProShop 三平台各编译验证一次（R64）。
  ------------------------------------------------------------------
  边界 Boundary     :
                      一 基准无效闸：dtIn 早于 DT#1970-01-01-00:00:00 视为未初始化或非法
                         时间戳，返回哨兵零点 + 信息级码 + bValid = FALSE，禁止把负天数
                         MOD 成一个看似合法的时刻（还原方向不饱和，R81：返回哨兵零点）；
                      二 日模 86400 显式化：diSecOfDay = ((纪元秒 MOD 86400) + 86400) MOD 86400，
                         双 MOD 保证负数路径也不落到负值域（域外不可达，证明在注释内）；
                      三 todOut 经 FC_DL_DintMsToTod 还原（毫秒域 × 1000），不自行拼 TOD 位型；
                      四 委托件的返回值与 bValid 由两个独立变量承接（R62-D5 教训：禁双写）；
                      五 纯函数：无记忆量、无定时器、无边沿实例，每调用重算。
  错误码 Codes      :
    16#0001_0652【信息级】输入时刻早于纪元基准，已返哨兵零点（bValid = FALSE，不置 bError）
    委托件故障码（16#0001_0330 / 0331 等）按「码随属主」原样回传（R66），本件不另立码。
  码位反证 Note     :
    本件唯一自有码 0652 不可省略：「早于基准」与「委托件进位失败」在出口上都是 bValid = FALSE
    且 todOut = 零点，但两者的处置主体与责任方不同（调用方时间戳未初始化 vs 平台位型承载异常），
    合并会让现场把「未初始化」误判为平台缺陷（R90 反证句）。
  验收 Acceptance   :
    算法已证（脚本）：未跑 ｜ 编译器已证（三平台）：未跑
    V1 DT#1970-01-01-00:00:00 → 0 秒、todOut = 00:00:00、bValid = TRUE
    V2 DT#2024-02-29-23:59:59 → 86399 秒（闰日不计日差，只取当日秒）
    V3 DT#2024-03-01-00:00:00 → 0 秒（日推进不残留）
    V4 DT#1970-01-01-00:00:00 之前的时刻 → bValid = FALSE + 码 0652 + 哨兵零点
    V5 DT#2106-02-07-06:28:15 → 23295 秒（6×3600 + 28×60 + 15，当日秒，跨 32 位不溢出）
    V6 DT#1970-01-02-00:00:00 → 0 秒（日推进归零）
  修订记录 Revision  :
    2026-11-21  v1.0.0  R62 首版（批 3 · 序号 7）
  ==================================================================
*)
FUNCTION FC_DL_DtToTodWrap : BOOL
VAR_INPUT
    dtIn : DT := DT#1970-01-01-00:00:00; // 输入时刻 [日期时间]，有效域自 1970-01-01-00:00:00 起 / the input instant, the domain starts at the epoch
END_VAR
VAR_OUTPUT
    todOut     : TOD;   // 当日时刻 [时刻]，00:00:00 ~ 23:59:59 / the time of day
    diSecOfDay : DINT;  // 当日秒数 [秒]，0..86399 / the second of the day
    bValid     : BOOL;  // 输出可用（早于基准与委托故障为 FALSE）[-] / the output is usable
    eErr       : UDINT; // 错误码，0 = 正常 / the error code, zero is ok
    bError     : BOOL;  // 故障标志，故障级码同拍置位（R45 配对）；信息级恒 FALSE / the fault flag, raised with a fault level code only
END_VAR
VAR
    _nEpochSec   : DINT := 0;                // 委托返回的纪元秒 [秒] / the epoch second returned by the delegate
    _bEpochValid : BOOL := FALSE;            // 委托 bValid 承接量（独立承接，禁双写）/ the delegate valid holder, never double written
    _bEpochErr   : BOOL := FALSE;            // 委托 bError 承接量（独立承接）/ the delegate fault holder, never double written
    _uEpochErr   : UDINT := 16#0000_0000;    // 委托错误码承接量 [码] / the delegate error code holder
    _nMsOfDay    : DINT := 0;                // 当日毫秒偏移 [毫秒] / the millisecond offset inside the day
    _todWork     : TOD := TOD#00:00:00;      // 委托 TOD 返回值承接量 [时刻] / the delegate time of day holder
    _bTodValid   : BOOL := FALSE;            // 委托 TOD 可用位承接量 / the delegate time of day usable holder
    _bTodErr     : BOOL := FALSE;            // 委托 TOD 故障位承接量 / the delegate time of day fault holder
    _uTodErr     : UDINT := 16#0000_0000;    // 委托 TOD 错误码承接量 [码] / the delegate time of day error code holder
    _bTodClamped : BOOL := FALSE;            // 委托 TOD 钳位位承接量（仅留档，不参与分级）/ the delegate clamp holder, recorded only
END_VAR  // R64 结构补齐：VAR 段缺失的 END_VAR（门禁机械修复）
VAR CONSTANT
    DL_DTT_SEC_PER_DAY : DINT := 86400;      // 每日秒数（日模）[秒] / the seconds of one day, the day modulus
    DL_DTT_MS_PER_SEC : DINT := 1000;        // 每秒毫秒数（毫秒域换算）[毫秒] / the milliseconds of one second
    DL_DTT_DINT_ZERO : DINT := 0;             // 整型零常量 [秒] / the integer zero constant
    DL_DTT_TOD_ZERO : TOD := TOD#00:00:00;   // 时刻哨兵零点 [时刻] / the sentinel midnight
    DL_DTT_EPOCH : DT := DT#1970-01-01-00:00:00; // 纪元基准时刻 [日期时间] / the epoch baseline instant
END_VAR

// 段 1｜返回值与全部出口预置安全值（R45 四段式第一段）/ segment 1, preset every outlet to its safe value
FC_DL_DtToTodWrap := FALSE; // 返回值预置假 / preset the return false
todOut := DL_DTT_TOD_ZERO; // 时刻预置哨兵零点 [时刻] / preset the sentinel midnight
diSecOfDay := DL_DTT_DINT_ZERO; // 当日秒数预置零 [秒] / preset the second of the day zero
bValid := FALSE; // 可用标志预置假，过闸后置位 / preset the validity false, raised after the gates
eErr := 16#0000_0000; // 错误码预置正常 / preset the code to ok
bError := FALSE; // 故障标志预置假 / preset the fault flag false
_nEpochSec := DL_DTT_DINT_ZERO; // 纪元秒承接量清零 [秒] / clear the epoch second holder
_bEpochValid := FALSE; // 委托可用位承接量清零 / clear the delegate usable holder
_bEpochErr := FALSE; // 委托故障位承接量清零 / clear the delegate fault holder
_uEpochErr := 16#0000_0000; // 委托码承接量清零 [码] / clear the delegate code holder
_nMsOfDay := DL_DTT_DINT_ZERO; // 当日毫秒清零 [毫秒] / clear the millisecond offset
_todWork := DL_DTT_TOD_ZERO; // 时刻承接量清零 [时刻] / clear the time of day holder
_bTodValid := FALSE; // 委托 TOD 可用位清零 / clear the time of day usable holder
_bTodErr := FALSE; // 委托 TOD 故障位清零 / clear the time of day fault holder
_uTodErr := 16#0000_0000; // 委托 TOD 码清零 [码] / clear the time of day code
_bTodClamped := FALSE; // 委托钳位位清零 / clear the delegate clamp holder

// 段 2｜基准无效闸：早于纪元的时刻不交给委托件（边界一，还原方向不饱和，R81）/ segment 2, the epoch baseline gate
IF dtIn < DL_DTT_EPOCH THEN // 未初始化或非法时间戳 / an uninitialised or illegal timestamp
    todOut := DL_DTT_TOD_ZERO; // 哨兵零点 [时刻] / the sentinel midnight
    diSecOfDay := DL_DTT_DINT_ZERO; // 哨兵零秒 [秒] / the sentinel zero second
    bValid := FALSE; // 输出不可用 / the output is not usable
    eErr := 16#0001_0652; // 信息级：输入早于纪元基准 / informational, the input precedes the epoch baseline
    bError := FALSE; // 明确不置故障标志（信息级，R285）/ keep the fault flag false, this is informational
    RETURN; // 早退，绝不把负天数交给委托件 / early return, a negative day count never reaches the delegate
END_IF

// 段 3｜委托时刻→纪元秒（R140 委托优先；返回值与可用位分承）/ segment 3, delegate the instant to the epoch second
_nEpochSec := FC_DL_DtToDintEpoch(dtIn := dtIn, eErr => _uEpochErr, bError => _bEpochErr, bValid => _bEpochValid); // 委托纪元秒换算 [秒] / delegate the epoch conversion
IF (NOT _bEpochValid) OR _bEpochErr THEN // 委托失败：码随属主回传（R66）/ the delegate failed, the code follows its owner
    eErr := _uEpochErr; // 原样回传委托码 [码] / replay the delegate code as is
    bError := _bEpochErr; // 原样回传委托故障位 / replay the delegate fault bit as is
    bValid := FALSE; // 输出不可用 / the output is not usable
    todOut := DL_DTT_TOD_ZERO; // 哨兵零点 [时刻] / the sentinel midnight
    diSecOfDay := DL_DTT_DINT_ZERO; // 哨兵零秒 [秒] / the sentinel zero second
    RETURN; // 早退 / early return
END_IF

// 段 4｜日模 86400 抽取当日秒（边界二：双 MOD 保证任何输入都落 0..86399）/ segment 4, the day modulus extraction
// 域外不可达证明：段 2 已证 dtIn ≥ 纪元，委托件已证返回值非负，故首层 MOD 的结果已在 [0, 86399]；
// 第二次「+ 86400 再 MOD」为结构对称的二重防御，保证任何未来改动都不会引入负值域出口。
// domain proof: the gate above guarantees a non negative epoch second, so the first modulus already lands inside the day;
// the second fold is a structural second line of defence against any future refactor.
diSecOfDay := ((_nEpochSec MOD DL_DTT_SEC_PER_DAY) + DL_DTT_SEC_PER_DAY) MOD DL_DTT_SEC_PER_DAY; // 当日秒数 [秒] / the second of the day

// 段 5｜委托毫秒→TOD 还原（边界三：不自行拼 TOD 位型）/ segment 5, delegate the millisecond offset back to a time of day
_nMsOfDay := diSecOfDay * DL_DTT_MS_PER_SEC; // 当日毫秒偏移（上界 86399000，DINT 内不溢出）[毫秒] / the millisecond offset, bounded by eighty six million four hundred thousand
_todWork := FC_DL_DintMsToTod(nMsOfDay := _nMsOfDay, bClampSilently := TRUE, eErr => _uTodErr, bError => _bTodErr, bValid => _bTodValid, bClamped => _bTodClamped); // 委托还原 [时刻] / delegate the restoration
IF (NOT _bTodValid) OR _bTodErr THEN // 委托失败：码随属主回传 / the delegate failed, the code follows its owner
    eErr := _uTodErr; // 原样回传委托码 [码] / replay the delegate code as is
    bError := _bTodErr; // 原样回传委托故障位 / replay the delegate fault bit as is
    bValid := FALSE; // 输出不可用 / the output is not usable
    todOut := DL_DTT_TOD_ZERO; // 哨兵零点 [时刻] / the sentinel midnight
    RETURN; // 早退 / early return
END_IF

// 段 6｜统一出口 / segment 6, the unified outlet
todOut := _todWork; // 时刻出口 [时刻] / the time of day outlet
bValid := TRUE; // 域内输出可用 / the in-domain output is usable
FC_DL_DtToTodWrap := TRUE; // 返回成功 / return success
END_FUNCTION

(* ---- FC_DL_DwordToHexString.st ---- *)
(*
    组件名称 : FC_DL_DwordToHexString
    所属子库 : DL_MathData
    当前版本 : 1.0.0
    兼 容 性 : CODESYS V3.5+ / TwinCAT 3 / 汇川 InoProShop；仅依赖 Standard.library
    功能描述 : DWORD → 8 位定宽十六进制文本，是 FC_DL_HexStringToBytes 的逆向对偶。
              取舍 ①：禁委托平台 DWORD_TO_STRING 的进制参数 —— 三家平台对「是否有 16# 前缀」「大小写」
              「是否补前导零」「不足位是否加空格」四项行为各不相同，一条日志换个平台就变样，
              报文回放与时间戳对齐全崩。本件用半字节查表 + CONCAT 自建，输出形态完全确定。
              取舍 ②：必须保留前导零（8 位定宽）—— 定宽是日志列对齐、二进制报文逐字节比对的前提；
              可变的短形态看着干净，却让「按位置切列」的所有下游脚本失效。
              取舍 ③：结果长度做出口自证 —— 若调用方把返回值声明成过短的 STRING，平台会静默截断，
              得到「看着像十六进制、其实少了几位」的串；本件比对实际长度与期望长度，不等即判故障并返回全零串，
              绝不交出一个长度不对的十六进制文本。
    开源溯源 : 原创实现（T0-6 字符串化变体线，HexStringToBytes R9 的逆向件）。无外部源码参考，；本件为 IEC 61131-3 标准语义的道莅防御性实现（原创实现，零外部源码复制）。
              码位与分级 100% 自有。预留槽说明：纯格式化函数的故障域天然窄，038E/038F/044A/044B
              为后续 bPadZero = FALSE（非定宽变体）保留，本轮实现体内零赋值。
    本文件内含 : FUNCTION FC_DL_DwordToHexString（单 POU，无配套类型）
    依 赖 : 无 DL_ 内部依赖；Standard.library: LEN / MID / CONCAT
    红线自检 : R1 ✓ 零全局变量与外部变量 ｜ R2 ✓ 零物理 IO 地址
              R3 ✓ 纯 IEC 61131-3 ｜ R4 ✓ 移位量恒 < 32（nIdx × 4 ≤ 28）+ 半字节掩码 + 出口长度自证
              R5 ✓ 全变量中英双语同行注释 ｜ R6 N/A 纯函数无顺序状态机，无 CASE 可写
              R7 N/A 无定时器、无沿检测实例 ｜ R8 ✓ 位数、半字节掩码、表串、前缀长度全常量化
    错误码   : 16#0001_044A [信息级] 预留禁用（不得挪用，留给 bPadZero = FALSE 变体）
               16#0001_044B [信息级] 预留禁用（不得挪用）
               16#0001_038D [故障级] 结果长度与期望不符（目标串长不足已被平台截断），返回 '00000000'，bValid = FALSE
               16#0001_038E [故障级] 预留禁用（不得挪用）
               16#0001_038F [故障级] 预留禁用（不得挪用）
    码位总账 : 16#0001_044A 预留 / 16#0001_044B 预留 ｜ 16#0001_038D 用 / 16#0001_038E 预留 / 16#0001_038F 预留
    遗留假设 : ① 返回类型声明为 STRING（平台缺省长度的具体值未知，CODESYS 缺省 80、部分平台缺省 256）；
              本件不假设长度，改用出口自证兜住。该自证只能发现「已截断」，不能预防截断，属可观测性而非免疫。
              ② MID 参数序按 IEC 标准 MID(串, 长度, 位置)，与库内既有 9 处用法同序；平台差异需在编译门槛核对。
    修订历史 :
        2026-11-16  v1.0.0  首版，R21 批次 3 入库
*)
FUNCTION FC_DL_DwordToHexString : STRING
VAR_INPUT
    uValue          : DWORD;          // 待格式化的双字，全 32 位有效 [位图] / double word to format, all 32 bits are significant [bitmap]
    bUpperCase      : BOOL := TRUE;   // TRUE 输出大写 A~F，FALSE 输出小写 a~f / TRUE emits upper case hex digits, FALSE emits lower case
    bPrefix         : BOOL := FALSE;  // TRUE 输出 16# 前缀（结果长 11）/ TRUE emits the 16# prefix, making the result eleven characters long
END_VAR
VAR_OUTPUT
    eErr            : UDINT;          // 错误码，0=正常；16#0001_04XX 信息级 / 16#0001_03XX 故障级 / error id, 0=ok
    bError          : BOOL;           // 故障级标志，eErr 落 16#0001_03XX 时为 TRUE / fault flag, TRUE on fault-level eErr
    bValid          : BOOL;           // 返回值是否可用 / result usable flag
    nLength         : INT;            // 结果串的实际长度 [字符] / actual length of the result string [char]
END_VAR
VAR
    sRet            : STRING;         // 结果装配缓冲 [字符] / result assembly buffer [char]
    nNib            : INT;            // 当前半字节值 0~15 [无量纲] / current nibble value, 0..15 [dimensionless]
    nIdx            : INT;            // 半字节游标 7~0（高位在前）[无量纲] / nibble cursor from seven down to zero, most significant first [dimensionless]
    nJ              : INT;            // 升序循环变量（镜像下标用）[无量纲] / ascending loop var for mirrored index [dimensionless]
    nExpLen         : INT;            // 期望结果长度 [字符] / expected result length [char]
END_VAR
VAR CONSTANT
    DL_HEX_UPPER        : STRING := '0123456789ABCDEF';   // 大写半字节表，位置 1 起对应值 0~15 [字符] / upper case nibble table indexed from one [char]
    DL_HEX_LOWER        : STRING := '0123456789abcdef';   // 小写半字节表，位置 1 起对应值 0~15 [字符] / lower case nibble table indexed from one [char]
    DL_HEX_PREFIX       : STRING := '16#';                // 十六进制前缀（可选）/ optional hexadecimal prefix
    DL_HEX_DIGITS       : INT := 8;                       // 定宽位数，DWORD 恰 8 个半字节 [位] / fixed width, a DWORD has eight nibbles [digit]
    DL_HEX_NIB_BITS     : INT := 4;                       // 半字节位宽，移位量 = 游标 × 4 ≤ 28 [位] / nibble width, the shift never exceeds twenty eight [bit]
    DL_HEX_PREFIX_LEN   : INT := 3;                       // 前缀长度 [字符] / prefix length [char]
    DL_HEX_NIB_MASK     : DWORD := 16#0000_000F;          // 半字节掩码 [位图] / nibble mask [bitmap]
    DL_HEX_ONE          : INT := 1;                       // 单位哨兵，MID 位置 1 基 [无量纲] / unity sentinel, MID is one based [dimensionless]
    DL_HEX_FALLBACK     : STRING := '00000000';           // 故障回退串，长度恒为 8 [字符] / fault fallback text with a constant length of eight [char]
    DL_DWORD_ZERO       : DWORD := 16#0000_0000;          // 零哨兵 [位图] / zero sentinel [bitmap]
    DL_ERR_NONE         : UDINT := 16#0000_0000;          // 无故障 / no error
END_VAR

// 段 1｜返回值与错误状态预置 / segment 1, preset the return value and the error state
FC_DL_DwordToHexString := DL_HEX_FALLBACK;   // 故障缺省返回全零串 / fault default returns eight zeros
eErr    := DL_ERR_NONE;                      // 预置无错误 / preset no error
bError  := FALSE;                            // 预置无故障 / preset no fault
bValid  := FALSE;                            // 预置结果不可用 / preset unusable
nLength := 0;                                // 预置长度 0 / preset the length to zero
sRet    := '';                               // 缓冲清空 / clear the buffer

// 段 2｜可选的十六进制前缀 / segment 2, optional hexadecimal prefix
IF bPrefix THEN
    sRet := DL_HEX_PREFIX;                   // 前缀先入，保证定宽位数在后 / the prefix comes first so the fixed width digits follow it
END_IF

// 段 3｜逐半字节装配：高位在前，移位量 = 游标 × 4，最大 28 < 32 / segment 3, nibble assembly, the shift never reaches the container width
FOR nJ := 0 TO (DL_HEX_DIGITS - DL_HEX_ONE) DO
    nIdx := (DL_HEX_DIGITS - DL_HEX_ONE) - nJ;   // 镜像下标：R509 禁 DOWNTO / mirrored index, DOWNTO unsupported
    nNib := DWORD_TO_INT(SHR(uValue, nIdx * DL_HEX_NIB_BITS) AND DL_HEX_NIB_MASK);   // 取当前半字节 / extract the current nibble
    IF bUpperCase THEN
        sRet := CONCAT(sRet, MID(DL_HEX_UPPER, DL_HEX_ONE, nNib + DL_HEX_ONE));      // 大写表查字符 / look the digit up in the upper case table
    ELSE
        sRet := CONCAT(sRet, MID(DL_HEX_LOWER, DL_HEX_ONE, nNib + DL_HEX_ONE));      // 小写表查字符 / look the digit up in the lower case table
    END_IF
END_FOR

// 段 4｜出口长度自证：平台静默截断必须被发现 / segment 4, length self proof catches a silent platform truncation
nLength := LEN(sRet);                        // 实际长度 / the actual length
nExpLen := DL_HEX_DIGITS;                    // 期望长度先取 8 / the expected length starts at eight
IF bPrefix THEN
    nExpLen := nExpLen + DL_HEX_PREFIX_LEN;  // 带前缀时 11 / eleven with the prefix
END_IF
IF nLength <> nExpLen THEN
    FC_DL_DwordToHexString := DL_HEX_FALLBACK;   // 回退到定宽全零串，长度可预测 / fall back to a fixed width zero text
    eErr   := 16#0001_038D;                  // 目标串长不足（故障级）/ the target string is too short, fault level
    bError := TRUE;                          // 置故障标志 / raise the fault flag
    nLength := LEN(DL_HEX_FALLBACK);         // 对外长度与回退串一致 / report the fallback length
    RETURN;                                  // bValid 保持 FALSE / bValid stays FALSE
END_IF

// 段 5｜出口 / segment 5, exit
FC_DL_DwordToHexString := sRet;              // 输出定宽十六进制文本 / publish the fixed width hexadecimal text
bValid := TRUE;                              // 结果可用 / the result is usable
END_FUNCTION

(* ---- FC_DL_DwordToIntSat.st ---- *)
(*
    FC_DL_DwordToIntSat —— DWORD 到 INT 的降位饱和
    ------------------------------------------------------------------
    分类      : DL_MathData / Convert
    前缀      : FC_DL_
    版本      : 1.0.0
    溯源      : IEC 61131-3 标准语义的道莅防御性实现（DWORD 32 位无符号 → INT 16 位有符号）；
                域内委托平台内建 DWORD_TO_INT，本件不重实现数学内核；
                上饱和出口、无损模式复核、错误分级与码位 100% 自有；
                clean-room 重写，未复制任何闭源厂商源码，参考实现仅限 MIT/Apache 许可
    平台      : 纯 IEC 61131-3，CODESYS V3.5+ / TwinCAT 3 / InoProShop 通用
    作者      : 道莅代码库 · PLC编程专家（R20）
    ------------------------------------------------------------------
    功能说明  : 长计数器、累计电量、批次总数这类 32 位累计值往 16 位 HMI 或老表写时，
                必须显式降位：本件统一取上饱和口径（钳到 32767），不做截断、不做回绕。
                截断会让 HMI 显示成随机跳动的小数，比钳位危险得多。
                核心防御：① 比较一律在 DWORD 字面量常量之间进行，绝不把 INT 上限先当 INT
                   再与 DWORD 比（隐式跨符号域比较在平台间有歧义，R56 纪律）；
                ② 上饱和置 bSatHigh 供 HMI 显示「已封顶」，避免把 32767 误读成真实值；
                ③ bRequireLossless = TRUE 时任何饱和即升故障级——结算与报表场景
                   不容许静默封顶，宁可停机也不出错数；
                ④ 域内路径零钳位、零额外比较开销。
                职责边界：WORD 16 位双语义归 FC_DL_WordToIntSat（它有补码口径），
                LWORD 64 位降位归 FC_DL_LwordToLintSat；本件只管 32 → 16 上饱和。
    编译门槛  : 主路径依赖平台内建 DWORD_TO_INT，IEC 61131-3 标准转换函数，
                三平台标准库均提供，无厂商方言。
    错误码    : 16#0001_0418 超域已饱和至 32767（bSatHigh 可查）——信息级，值可用
                16#0001_0419 预留禁用（信息级，不得挪用）
                16#0001_0342 调用方要求无损（bRequireLossless = TRUE）却发生饱和——故障级，bValid = FALSE
                16#0001_0343 预留（故障级，不得挪用）
                16#0001_0344 预留禁用（故障级，不得挪用）
    码位总账  : 16#0001_0418 用 / 16#0001_0419 预留 ｜ 16#0001_0342 用 / 16#0001_0343 预留 / 16#0001_0344 预留
    状态机    : R6 标注 N/A —— 本组件为纯函数无顺序状态机，无 CASE 可写，非法状态不可能出现
    采样约定  : 本件无定时器、无沿检测、无状态；单拍纯计算，结论与任务周期无关。
    修订记录  : 2026-11-16 v1.0.0 首次入库（R20）
*)
FUNCTION FC_DL_DwordToIntSat : INT
VAR_INPUT
    uIn              : DWORD;                 // 输入值 [无量纲]，全域 0~4294967295 / input value [dimensionless], full DWORD domain
    bRequireLossless : BOOL := FALSE;         // TRUE = 发生饱和即判故障（计量/结算场景）/ TRUE turns any saturation into a fault
END_VAR
VAR_OUTPUT
    eErr             : UDINT;                 // 错误码，0=正常 / error id, 0=ok
    bError           : BOOL;                  // 故障标志，eErr 为故障级时 TRUE / error flag, TRUE on fault-level eErr
    bValid           : BOOL;                  // 返回值是否可用（要求无损却饱和时为 FALSE）/ return usable, FALSE when saturated in lossless mode
    bSatHigh         : BOOL;                  // 上饱和发生（输入 > 32767）/ high saturation occurred
END_VAR
VAR CONSTANT
    DL_INT_MAX_AS_DWORD : DWORD := 32767;     // INT 上限的 DWORD 形态 [无量纲] / the INT maximum expressed as DWORD [dimensionless]
    DL_INT_MAX       : INT := 32767;          // INT 上限值 [无量纲] / the INT maximum value [dimensionless]
    DL_INT_ZERO      : INT := 0;              // 有符号零常量，避免裸字面量 [无量纲] / signed zero constant [dimensionless]
END_VAR
VAR
    nOut             : INT;                   // 结果中间量 [无量纲] / result intermediate [dimensionless]
END_VAR

// 段 1｜返回值与错误状态预置 / segment 1, preset return value and error status
FC_DL_DwordToIntSat := DL_INT_ZERO;           // 故障缺省返回 0 [无量纲] / fault default returns zero [dimensionless]
eErr := 0;                                    // 预置无错误 / preset no error
bError := FALSE;                              // 预置无故障 / preset no fault
bValid := FALSE;                              // 预置不可用，通过闸门后置位 / preset invalid, set TRUE after the gates
bSatHigh := FALSE;                            // 预置未饱和 / preset no saturation
nOut := DL_INT_ZERO;                          // 结果中间量清零 / clear the result intermediate

// 段 2｜降位闸：用 DWORD 字面量比较，禁跨符号域比较 / segment 2, narrowing gate with a DWORD literal comparison
IF uIn > DL_INT_MAX_AS_DWORD THEN
    nOut := DL_INT_MAX;                       // 上饱和至 32767 / saturate to the INT maximum
    bSatHigh := TRUE;                         // 标记上饱和 / flag the high saturation
    eErr := 16#0001_0418;                     // 信息级：超域已饱和 / info level, saturated on the overrun
ELSE
    // 段 3｜域内才委托内建 / segment 3, delegate only inside the domain
    nOut := DWORD_TO_INT(uIn);                // 域内无损降位 [无量纲] / lossless narrowing inside the domain [dimensionless]
END_IF

// 段 4｜无损模式复核（要求无损却发生饱和即故障级）/ segment 4, lossless recheck
IF bRequireLossless AND bSatHigh THEN
    eErr := 16#0001_0342;                     // 故障级：要求无损却发生饱和 / fault level, saturation under the lossless requirement
    bError := TRUE;                           // 置故障标志 / raise the error flag
    bValid := FALSE;                          // 返回值不可进结算 / the value must not enter settlements
    FC_DL_DwordToIntSat := nOut;              // 仍发布钳位值供 HMI 观察 / still publish the clamped value for observation
    RETURN;                                   // 出口 / exit
END_IF

// 段 5｜发布结果 / segment 5, publish the result
FC_DL_DwordToIntSat := nOut;                  // 输出 16 位有符号结果 [无量纲] / publish the signed 16-bit result [dimensionless]
bValid := TRUE;                               // 直通或钳位均可用 / usable either way
bError := FALSE;                              // 信息级不置故障 / info level never raises a fault
END_FUNCTION

(* ---- FC_DL_ElectrolyzerCellVoltageCalc.st ---- *)
(*
  DL Factory R88 | FC_DL_ElectrolyzerCellVoltageCalc
  功能：工程简化单槽电压 U=U_rev+R·i+s·ln(i/i0)（可逆电压+欧姆+塔菲尔），超 2.0 V 报警
  开源溯源：无（clean-room 自研，依据公开工艺公式 电解槽电压分解式 U=U_rev+iR+η_act，许可证=MIT，借鉴点=公式结构）
  规则：R1-R16 全遵守；R88 简单件标量形（纯标量入参出参，无循环体、无方法、无属性、无数组）
*)
FUNCTION FC_DL_ElectrolyzerCellVoltageCalc : REAL
VAR_INPUT
    fUrevV : REAL := 1.23; // 可逆（热中性参考）电压 U_rev @25°C [V] / reversible voltage [V]
    fRohmOhmCm2 : REAL := 0.15; // 面积比欧姆电阻（含膜与接触） [Ω·cm²] / area specific ohmic resistance [ohm*cm^2]
    fCurrentDensityAPerCm2 : REAL := 0.5; // 电流密度 i [A/cm²] / current density [A/cm^2]
    fTafelSlopeV : REAL := 0.05; // 塔菲尔斜率 s（每数量级电压增量） [V/dec] / tafel slope [V/dec]
    fExchangeCurrentDensityAPerCm2 : REAL := 1.0E-3; // 交换电流密度 i0（ln 的基准） [A/cm²] / exchange current density [A/cm^2]
    fLimitV : REAL := 2.0; // 单槽电压报警上限（能效恶化提示） [V] / cell voltage alarm limit [V]
END_VAR
VAR_OUTPUT
    fCellV : REAL; // 单槽电压 U [V] / cell voltage [V]
    xOverLimit : BOOL; // TRUE=单槽电压超过报警上限 [-] / TRUE when above the alarm limit [-]
END_VAR
VAR
    fRatio : REAL; // i/i0（对数量纲一化比值） [-] / current density ratio [-]
    fOhmicV : REAL; // 欧姆压降 i·R [V] / ohmic drop [V]
    fActV : REAL; // 活化过电位 s·ln(i/i0) [V] / activation overpotential [V]
END_VAR

// 段 1｜出口预置
FC_DL_ElectrolyzerCellVoltageCalc := -1.0; // 哨兵返回 -1（无效） [-] / sentinel return -1, invalid [-]
fCellV := 0.0; // 单槽电压预置零 [V] / cell voltage preset zero [V]
xOverLimit := FALSE; // 超限位预置 FALSE（未判定前不报警） [-] / over-limit flag preset false [-]

// 段 2｜非有限拦截 + 域闸
IF NOT (fUrevV > -1.0E30 AND fUrevV < 1.0E30) OR NOT (fRohmOhmCm2 > -1.0E30 AND fRohmOhmCm2 < 1.0E30) OR NOT (fCurrentDensityAPerCm2 > -1.0E30 AND fCurrentDensityAPerCm2 < 1.0E30) THEN
    RETURN; // 可逆电压/欧姆电阻/电流密度任一非有限即拒算 [-] / any non finite input rejected [-]
END_IF
IF NOT (fTafelSlopeV > -1.0E30 AND fTafelSlopeV < 1.0E30) OR NOT (fExchangeCurrentDensityAPerCm2 > -1.0E30 AND fExchangeCurrentDensityAPerCm2 < 1.0E30) OR NOT (fLimitV > -1.0E30 AND fLimitV < 1.0E30) THEN
    RETURN; // 塔菲尔斜率/i0/上限任一非有限则判据静默失效，故先拦 [-] / these pins must be finite [-]
END_IF
IF fCurrentDensityAPerCm2 < 1.0E-9 OR fExchangeCurrentDensityAPerCm2 < 1.0E-9 THEN
    RETURN; // ln 的自变量须为正：i 与 i0 都必须大于 1E-9 [A/cm²] / ln argument must be positive [A/cm^2]
END_IF
IF fRohmOhmCm2 < 0.0 OR fTafelSlopeV < 0.0 OR fUrevV <= 0.0 OR fLimitV <= 0.0 THEN
    RETURN; // 物理符号域闸：电阻/斜率非负、可逆电压与上限为正 [Ω·cm², V] / physical sign gates [-]
END_IF

// 段 3｜计算
fRatio := fCurrentDensityAPerCm2 / fExchangeCurrentDensityAPerCm2; // (A/cm²) ÷ (A/cm²) = 无量纲 [-] / dimensionless ratio [-]
IF fRatio < 1.0E-9 THEN
    RETURN; // 除法后复核：比值须为正，否则 LN 产生非有限值 [-] / ratio must stay positive before LN [-]
END_IF
fOhmicV := fRohmOhmCm2 * fCurrentDensityAPerCm2; // (Ω·cm²) × (A/cm²) = V，量纲自洽 [V] / [ohm*cm^2] x [A/cm^2] = [V]
fActV := fTafelSlopeV * LN(fRatio); // V × 无量纲 = V，活化过电位 [V] / [V] x [-] = [V]
fCellV := fUrevV + fOhmicV + fActV; // V + V + V = V，三项分解合成 [V] / [V]

// 段 4｜判定与饱和
IF NOT (fCellV > -1.0E30 AND fCellV < 1.0E30) THEN
    RETURN; // 结果非有限再拦一次 [-] / re-check the result for finiteness [-]
END_IF
xOverLimit := fCellV > fLimitV; // 严格大于上限为报警，等于上限仍判正常 [V] / strict compare [V]

// 段 5｜出口自检
IF fCellV < fUrevV THEN
    RETURN; // 出口自检：单槽电压不应低于可逆电压（过电位恒非负） [V] / cell voltage must not drop below U_rev [V]
END_IF
FC_DL_ElectrolyzerCellVoltageCalc := fCellV; // 返回单槽电压 U [V] / return the cell voltage [V]
END_FUNCTION

(* ---- FC_DL_ElectrolyzerH2RateCalc.st ---- *)
(*
  DL Factory R88 | FC_DL_ElectrolyzerH2RateCalc
  功能：法拉第定律算电解槽产氢体积流量 V_H2=n·I·η_F/(2F)·Vm，并给出电流密度（按单槽活性面积）
  开源溯源：无（clean-room 自研，依据公开工艺公式 法拉第电解定律 V=n·I·η/(2F)·Vm，许可证=MIT，借鉴点=公式结构）
  规则：R1-R16 全遵守；R88 简单件标量形（纯标量入参出参，无循环体、无方法、无属性、无数组）
*)
FUNCTION FC_DL_ElectrolyzerH2RateCalc : REAL
VAR_INPUT
    fCurrentA : REAL := 10000.0; // 电解电源电流 I（整堆串联电流，各槽相同） [A] / stack current [A]
    fCells : REAL := 100.0; // 串联电解槽（单胞）数量 n [个] / number of series cells [-]
    fFaradEff : REAL := 0.98; // 法拉第效率 η_F（0~1，含气体交叉损失） [-] / faradaic efficiency [-]
    fCellAreaCm2 : REAL := 1000.0; // 单槽活性面积 A [cm²] / single cell active area [cm^2]
END_VAR
VAR_OUTPUT
    fH2Nm3h : REAL; // 标准状态产氢体积流量 [Nm³/h] / hydrogen flow at standard conditions [Nm^3/h]
    fCurrentDensityAPerCm2 : REAL; // 电流密度 i=I/A [A/cm²] / current density [A/cm^2]
END_VAR
VAR
    fFaradayC : REAL; // 法拉第常数 F（库仑/摩尔电子） [C/mol] / faraday constant [C/mol]
    fTwoF : REAL; // 分母 2F（每摩尔 H2 需 2 mol 电子） [C/mol] / the 2F divisor [C/mol]
    fMolPerS : REAL; // 产氢摩尔流率 [mol/s] / hydrogen molar flow [mol/s]
END_VAR

// 段 1｜出口预置
FC_DL_ElectrolyzerH2RateCalc := -1.0; // 哨兵返回 -1（无效） [-] / sentinel return -1, invalid [-]
fH2Nm3h := 0.0; // 产氢流量预置零 [Nm³/h] / hydrogen flow preset zero [Nm^3/h]
fCurrentDensityAPerCm2 := 0.0; // 电流密度预置零 [A/cm²] / current density preset zero [A/cm^2]

// 段 2｜非有限拦截 + 域闸
IF NOT (fCurrentA > -1.0E30 AND fCurrentA < 1.0E30) OR NOT (fCells > -1.0E30 AND fCells < 1.0E30) THEN
    RETURN; // 电流/槽数任一非有限即拒算 [-] / any non finite input rejected [-]
END_IF
IF NOT (fFaradEff > -1.0E30 AND fFaradEff < 1.0E30) OR NOT (fCellAreaCm2 > -1.0E30 AND fCellAreaCm2 < 1.0E30) THEN
    RETURN; // 法拉第效率/活性面积任一非有限即拒算 [-] / any non finite input rejected [-]
END_IF
IF fCurrentA < 0.0 OR fCells < 1.0 THEN
    RETURN; // 电流非负闸 + 槽数下限闸（整数语义，至少 1 个单胞） [A, 个] / non negative current and one cell at least
END_IF
IF fFaradEff <= 0.0 OR fFaradEff > 1.0 OR fCellAreaCm2 < 1.0E-9 THEN
    RETURN; // 法拉第效率开区间闸 (0,1] + 活性面积正域闸（面积是分母） [-] / efficiency and area gates
END_IF

// 段 3｜计算（A→mol/s→Nm³/h 链路，逐项量纲见行尾注释）
fFaradayC := 96485.0; // 法拉第常数装入 [C/mol] / load the faraday constant [C/mol]
fTwoF := 2.0 * fFaradayC; // 2 × C/mol = C/mol，每摩 H2 需 2 摩电子 [C/mol] / [C/mol]
IF fTwoF < 1.0E-9 THEN
    RETURN; // 除法前分母闸：2F 必须大于 1E-9 才可作除数 [C/mol] / denominator gate [C/mol]
END_IF
fMolPerS := fCurrentA * fCells * fFaradEff / fTwoF; // A × 个 × 无量纲 ÷ (C/mol) = mol/s，法拉第定律 [mol/s] / [mol/s]
fH2Nm3h := fMolPerS * 22.414 * 3600.0 * 0.001; // (mol/s) × 22.414 L/mol × 3600 s/h × 0.001 m³/L = Nm³/h [Nm³/h] / [Nm^3/h]
IF fCellAreaCm2 < 1.0E-9 THEN
    RETURN; // 除法前分母闸：活性面积必须大于 1E-9 才可作除数 [cm²] / denominator gate [cm^2]
END_IF
fCurrentDensityAPerCm2 := fCurrentA / fCellAreaCm2; // A ÷ cm² = A/cm²，电流密度 [A/cm²] / [A/cm^2]

// 段 4｜判定与饱和
IF NOT (fH2Nm3h > -1.0E30 AND fH2Nm3h < 1.0E30) OR NOT (fCurrentDensityAPerCm2 > -1.0E30 AND fCurrentDensityAPerCm2 < 1.0E30) THEN
    RETURN; // 两出口非有限再拦一次 [-] / re-check both results for finiteness [-]
END_IF

// 段 5｜出口自检
IF fH2Nm3h < 0.0 THEN
    RETURN; // 出口自检：产氢流量不得为负（负值说明电流符号错） [Nm³/h] / flow must not be negative [Nm^3/h]
END_IF
FC_DL_ElectrolyzerH2RateCalc := fH2Nm3h; // 返回标准状态产氢体积流量 [Nm³/h] / return the hydrogen flow [Nm^3/h]
END_FUNCTION

(* ---- FC_DL_ElectrolyzerKohConcCalc.st ---- *)
(*
  DL Factory R88 | FC_DL_ElectrolyzerKohConcCalc
  功能：由碱液密度反算 KOH 质量分数 w%=(ρ-1.0)/0.0105，并给经验电导率估计（线性经验式）
  开源溯源：无（clean-room 自研，依据公开工艺公式 碱液密度-浓度线性近似与电导率经验式，许可证=MIT，借鉴点=公式结构）
  规则：R1-R16 全遵守；R88 简单件标量形（纯标量入参出参，无循环体、无方法、无属性、无数组）
*)
FUNCTION FC_DL_ElectrolyzerKohConcCalc : REAL
VAR_INPUT
    fDensityGcm3 : REAL := 1.28; // 碱液密度 ρ（20~25°C 实测） [g/cm³] / electrolyte density [g/cm^3]
    fSlopeGcm3PerPct : REAL := 0.0105; // 密度对质量分数的经验斜率（每 1% 浓度） [g/cm³/%] / empirical density slope [g/cm^3 per pct]
    fCondCoeffSPerCm : REAL := 0.02; // 电导率经验系数（满量程前置系数） [S/cm] / empirical conductivity coefficient [S/cm]
END_VAR
VAR_OUTPUT
    fMassPct : REAL; // KOH 质量分数 w [%] / KOH mass fraction [%]
    fCondSPerCm : REAL; // 电导率经验估计 σ [S/cm] / estimated conductivity [S/cm]
END_VAR
VAR
    fSlope : REAL; // 斜率缓存（除零判据） [g/cm³/%] / cached slope, the divisor [g/cm^3 per pct]
    fNetDensity : REAL; // 密度超出水的部分 ρ-1.0 [g/cm³] / density above that of water [g/cm^3]
END_VAR

// 段 1｜出口预置
FC_DL_ElectrolyzerKohConcCalc := -1.0; // 哨兵返回 -1（无效） [-] / sentinel return -1, invalid [-]
fMassPct := 0.0; // 质量分数预置零 [%] / mass fraction preset zero [%]
fCondSPerCm := 0.0; // 电导率预置零 [S/cm] / conductivity preset zero [S/cm]
fSlope := 0.0; // 斜率缓存预置零 [g/cm³/%] / slope preset zero [g/cm^3 per pct]
fNetDensity := 0.0; // 密度余量预置零 [g/cm³] / density surplus preset zero [g/cm^3]

// 段 2｜非有限拦截 + 域闸
IF NOT (fDensityGcm3 > -1.0E30 AND fDensityGcm3 < 1.0E30) OR NOT (fSlopeGcm3PerPct > -1.0E30 AND fSlopeGcm3PerPct < 1.0E30) THEN
    RETURN; // 密度/斜率任一非有限即拒算 [-] / any non finite input rejected [-]
END_IF
IF NOT (fCondCoeffSPerCm > -1.0E30 AND fCondCoeffSPerCm < 1.0E30) THEN
    RETURN; // 电导系数非有限则第二出口无意义，故先拦 [S/cm] / the coefficient must be finite [S/cm]
END_IF
IF fDensityGcm3 <= 1.0 OR fDensityGcm3 >= 1.35 THEN
    RETURN; // 密度开区间域闸 (1.0,1.35)：低于水或超饱和则线性近似失效 [g/cm³] / density open interval gate [g/cm^3]
END_IF
IF fSlopeGcm3PerPct < 1.0E-9 THEN
    RETURN; // 除法前分母闸：斜率必须大于 1E-9（同时为正域闸） [g/cm³/%] / denominator gate [g/cm^3 per pct]
END_IF
IF fCondCoeffSPerCm <= 0.0 THEN
    RETURN; // 电导系数正域闸：非正值会使第二出口恒零 [S/cm] / positive coefficient gate [S/cm]
END_IF

// 段 3｜计算（经验式：非标准定义，仅用于 25°C 附近粗估）
fSlope := fSlopeGcm3PerPct; // 取斜率作除数缓存 [g/cm³/%] / cache the slope as divisor [g/cm^3 per pct]
fNetDensity := fDensityGcm3 - 1.0; // g/cm³ - g/cm³ = g/cm³，扣掉水的密度 [g/cm³] / density above water [g/cm^3]
fMassPct := fNetDensity / fSlope; // (g/cm³) ÷ (g/cm³/%) = %，线性近似反算浓度 [%] / [g/cm^3] / [g/cm^3 per pct] = [%]
IF fMassPct <= 0.0 OR fMassPct >= 100.0 THEN
    RETURN; // 浓度开区间闸 (0,100)：反算越界说明线性近似不适用 [%] / open interval gate on the fraction [%]
END_IF
fCondSPerCm := fCondCoeffSPerCm * fMassPct * (1.0 - fMassPct * 0.01); // S/cm × % × 无量纲 = S/cm，抛物线型经验式 [S/cm] / [S/cm]

// 段 4｜判定与饱和
IF NOT (fMassPct > -1.0E30 AND fMassPct < 1.0E30) OR NOT (fCondSPerCm > -1.0E30 AND fCondSPerCm < 1.0E30) THEN
    RETURN; // 两出口非有限再拦一次 [-] / re-check both results for finiteness [-]
END_IF

// 段 5｜出口自检
IF fCondSPerCm <= 0.0 THEN
    RETURN; // 出口自检：电导率须为正，否则经验式参数被误用 [S/cm] / conductivity must be positive [S/cm]
END_IF
FC_DL_ElectrolyzerKohConcCalc := fMassPct; // 返回 KOH 质量分数 [%] / return the KOH mass fraction [%]
END_FUNCTION
